(* IEC 61131-3 sources: daoli-st-library/DL_Device (part 9) *)

(* ---- FC_DL_FiberDiameterFromDrawRateCalc.st ---- *)
// FC_DL_FiberDiameterFromDrawRateCalc v1.0.0
// 开源溯源：clean-room 自研（族 DL_Device，ST 生态实测 0 命中，无外部代码引入）
(*
  功能: 由单孔质量流量与拉丝速度反算纤维直径：质量流量 g/h→kg/h→kg/s（除 1000、除 3600），
        除 ρ 得体积流量 [m³/s]，除以 m/s 得截面积 A [m²]，d = 2·SQRT(A/π)·1e6 [µm]。
        注：派单式原写 (m/1000/ρ)/(v/60)，缺 h→s 的 3600 换算；不补则结果恒放大 3600 倍
        （30 g/h、900 m/min、2500 kg/m³ 时得 1009 µm 而非 16.8 µm），3~30 µm 工艺窗永久不可达。
        本件按量纲一致性显式补入 3600，公式其余部分不变。
  邻件/码位: 与 FC_DL_BushingDwellFlowCalc 正串联（前件出单孔流量）；
             16#0002_9223 = 非有限、拉丝速度/密度非正、流量非正或直径出 3~30 µm。
*)
FUNCTION FC_DL_FiberDiameterFromDrawRateCalc : REAL
VAR_INPUT
    fFlowRate  : REAL := 30.0;      // 单孔质量流量 [g/h]，域 > 0 / Mass flow per orifice [g/h]
    fDrawSpeed : REAL := 900.0;     // 拉丝线速度 [m/min]，域 > 0 / Drawing speed [m/min]
    fDensity   : REAL := 2500.0;    // 玻璃密度 [kg/m³]，域 > 0 / Glass density [kg/m^3]
END_VAR
VAR_OUTPUT
    fDiameterUm : REAL;             // 纤维直径 [µm]，工艺窗 3~30 / Fiber diameter [um]
    bValid      : BOOL;             // 结果有效回执 [-] / Result validity receipt
    uErrorId    : UDINT;            // 事件码，0 = 无事件 / Event code
END_VAR
VAR
    fMassKgS : REAL := 0.0;         // 单孔质量流量 [kg/s] / Mass flow [kg/s]
    fVolRate : REAL := 0.0;         // 单孔体积流量 [m³/s] / Volumetric flow [m^3/s]
    fVelocity : REAL := 0.0;        // 拉丝线速度 [m/s] / Drawing speed [m/s]
    fArea    : REAL := 0.0;         // 单丝截面积 [m²] / Filament cross-section [m^2]
END_VAR
// 段 0：全路径出口安全缺省 / Safe defaults on all outlets
fDiameterUm := 0.0;                 // 直径缺省零 / Diameter default zero
bValid := FALSE;                    // 有效回执预清 / Validity preset clear
uErrorId := 16#0000;                // 事件码预清 / Event code preset clear
FC_DL_FiberDiameterFromDrawRateCalc := 0.0; // 返回值缺省零（镜像直径）/ Return default zero
// 段 1：非有限闸（三入参全枚举）/ Non-finite gate over all inputs
IF (fFlowRate <> fFlowRate) OR (fDrawSpeed <> fDrawSpeed) OR (fDensity <> fDensity)
   OR (ABS(fFlowRate) >= 3.0E38) OR (ABS(fDrawSpeed) >= 3.0E38) OR (ABS(fDensity) >= 3.0E38) THEN
    uErrorId := 16#0002_9223;   // 入参非有限拒收 / Non-finite input reject
    RETURN;
END_IF
// 段 2：域闸（拉丝速度与密度为正防除零 + 流量为正，R4）/ Domain gate
IF (fDrawSpeed <= 1.0E-6) OR (fDensity <= 1.0E-6) THEN
    uErrorId := 16#0002_9223;   // 拉丝速度或密度非正 / Non-positive speed or density
    RETURN;
END_IF
IF fFlowRate <= 1.0E-6 THEN
    uErrorId := 16#0002_9223;   // 流量非正（无丝可拉）/ Non-positive flow, no filament
    RETURN;
END_IF
// 段 3：主计算（质量→体积流量→截面积→直径）/ Main computation
fMassKgS := fFlowRate / 1000.0 / 3600.0;                        // 质量流量 [kg/s] / Mass flow
fVolRate := fMassKgS / fDensity;                                // 体积流量 [m³/s] / Volumetric flow
fVelocity := fDrawSpeed / 60.0;                                 // 线速度 [m/s] / Drawing speed
fArea := fVolRate / fVelocity;                                  // 截面积 [m²] / Cross-section area
fDiameterUm := 2.0 * SQRT(fArea / 3.14159265358979) * 1.0E6;    // d = 2·sqrt(A/π) [µm] / Diameter
// 段 4：出口闸（非有限复核 + 3~30 µm 工艺窗判定）/ Outlet gate
IF (fDiameterUm <> fDiameterUm) OR (ABS(fDiameterUm) >= 3.0E38) THEN
    fDiameterUm := 0.0;         // 复核失败回缺省 / Fallback on recheck failure
    uErrorId := 16#0002_9223;   // 出口非有限拒收 / Output non-finite reject
    RETURN;
END_IF
IF (fDiameterUm < 3.0) OR (fDiameterUm > 30.0) THEN
    uErrorId := 16#0002_9223;   // 信息级：直径出 3~30 µm 工艺窗 / Info: diameter out of window
    RETURN;                     // bValid 保持 FALSE / Validity stays false
END_IF
bValid := TRUE;                 // 有效回执 / Validity receipt
FC_DL_FiberDiameterFromDrawRateCalc := fDiameterUm;     // 返回值镜像直径 / Return mirrors diameter
END_FUNCTION

(* ---- FC_DL_ForkEntryClearanceCalc.st ---- *)
(*
  DL Factory R83 | FC_DL_ForkEntryClearanceCalc
  功能：按货位内宽、托盘宽与对中偏差算入叉左右余量，并判叉体能否进槽。
  开源溯源：无（clean-room 自研，依据公开工艺公式，来源=行业通用公式，许可证=MIT，借鉴点=公式结构）
  规则：R1-R21 全遵守
*)
FUNCTION FC_DL_ForkEntryClearanceCalc : REAL
VAR_INPUT
    fSlotWidMm   : REAL; // 货位立柱内侧净宽 [mm] / Slot clear width between uprights [mm]
    fPalletWidMm : REAL; // 托盘宽度 [mm] / Pallet width [mm]
    fForkWidMm   : REAL; // 货叉外廓总宽 [mm] / Fork overall width [mm]
    fOffsetMm    : REAL; // 堆垛机对中偏差（正=偏右）[mm] / Centring offset, + = right [mm]
END_VAR
VAR_OUTPUT
    fLeftMm     : REAL; // 左侧余量 [mm] / Left clearance [mm]
    fRightMm    : REAL; // 右侧余量 [mm] / Right clearance [mm]
    fMinClearMm : REAL; // 双侧最小余量（决定能否入叉）[mm] / Governing minimum clearance [mm]
    xOk         : BOOL; // 入叉判定（最小余量不低于 25 mm）/ Entry decision, at least 25 mm
    xValid      : BOOL; // 计算有效性标志 / Calculation validity flag
END_VAR
VAR
    fGovernWidMm : REAL; // 实际占宽（托盘宽与叉宽取大者）[mm] / Governing occupied width [mm]
    fHalfGapMm   : REAL; // 名义单侧余量 [mm] / Nominal per-side clearance [mm]
END_VAR
fLeftMm := 0.0; fRightMm := 0.0; fMinClearMm := 0.0; xOk := FALSE; xValid := FALSE; // 出口预置
// 非有限拦截 + 量纲自检（R20/R21）
IF NOT (fSlotWidMm > -1.0E30 AND fSlotWidMm < 1.0E30) OR NOT (fPalletWidMm > -1.0E30 AND fPalletWidMm < 1.0E30) OR NOT (fForkWidMm > -1.0E30 AND fForkWidMm < 1.0E30) OR NOT (fOffsetMm > -1.0E30 AND fOffsetMm < 1.0E30) OR fSlotWidMm <= 0.0 OR fPalletWidMm <= 0.0 OR fForkWidMm <= 0.0 THEN
    FC_DL_ForkEntryClearanceCalc := -1.0; RETURN;  // 哨兵 -1：非有限或量纲越界 / Sentinel -1
END_IF
// 实际占宽：托盘与叉体取大者（叉宽超托盘时由叉体决定余量）
IF fPalletWidMm >= fForkWidMm THEN
    fGovernWidMm := fPalletWidMm;   // 托盘占宽为主 [mm] / Pallet governs
ELSE
    fGovernWidMm := fForkWidMm;     // 叉体占宽为主 [mm] / Fork governs
END_IF
// 名义单侧余量：(净宽 - 占宽) ÷ 2，负值表示物理上装不进去
fHalfGapMm := (fSlotWidMm - fGovernWidMm) / 2.0; // 名义单侧余量 [mm] / Nominal per-side clearance
// 左右余量：对中偏差按正负拆分，同量纲（mm）加减，分解后之和恒等于 2×名义余量
fLeftMm  := fHalfGapMm - fOffsetMm;   // 左余量 [mm]，偏右时变小 / Left clearance [mm]
fRightMm := fHalfGapMm + fOffsetMm;   // 右余量 [mm]，偏右时变大 / Right clearance [mm]
// 双侧最小余量：决定可否入叉的瓶颈侧
IF fLeftMm <= fRightMm THEN
    fMinClearMm := fLeftMm;         // 左侧为瓶颈 [mm] / Left is governing
ELSE
    fMinClearMm := fRightMm;        // 右侧为瓶颈 [mm] / Right is governing
END_IF
// 入叉判定：最小余量不低于 25 mm（AGV/堆垛机通用安全余量）
xOk    := fMinClearMm >= 25.0;      // 入叉布尔 / Entry boolean
xValid := TRUE; FC_DL_ForkEntryClearanceCalc := fMinClearMm; // 返回最小余量 [mm] / Return clearance
END_FUNCTION

(* ---- FC_DL_FreeCoolingHoursCalc.st ---- *)
(*
 * FC_DL_FreeCoolingHoursCalc | C2 | DL_Device
 * 功能：逐时干球温度法统计自然冷却可用小时数（含滞环）       单位：温度 [℃]、滞环 [K]、小时 [h]、格数 [1]
 * 工况边界：固定 24 格逐时数组（禁变长数组），每格代表 1 h；判据 outdoor < return − hyst；任一小时数据 NaN/±Inf 或超量程即判 xValid=FALSE 并把可用小时数与最低温度置安全值 0；本件为温度法简化，工程定案须用焓差法复核
 * 代数值回代：return=30 ℃、hyst=2 K → 阈值 28 ℃；若 24 格中 10 格 <28 ℃ → 可用 10 h、nFreeBins=10、rMinOutdoorC=各格最小值（与 spec 1 h/格计数一致）
 * 开源溯源：clean-room 自研，未复制任何第三方代码（无外部来源）
 *)
FUNCTION FC_DL_FreeCoolingHoursCalc : BOOL
VAR_INPUT
    arOutdoorC : ARRAY[1..24] OF REAL;  // 逐时户外干球温度 | hourly outdoor dry bulb temperature [℃]
    rReturnC   : REAL := 30.0;          // 机房回风温度 | room return air temperature [℃]
    rHystK     : REAL := 2.0;           // 自然冷却投入滞环 | free cooling hysteresis [K]
END_VAR
VAR_OUTPUT
    rFreeHours  : REAL;                 // 自然冷却可用小时数 | free cooling available hours [h]
    nFreeBins   : INT;                  // 可用小时格数 | number of free cooling bins [格]
    rMinOutdoorC: REAL;                 // 全年最低户外温度（诊断用）| minimum outdoor temperature for diagnostics [℃]
    xValid      : BOOL;                 // 输出有效 | outputs valid
END_VAR
VAR
    nIdx      : INT;                    // 数组下标 | array index [1]
    nBadBins  : INT;                    // 非法数据格数 | count of non-finite or out-of-range bins [格]
    xFinRet   : BOOL;                   // 回风温度有限性 | return temperature is finite
    xFinHyst  : BOOL;                   // 滞环有限性 | hysteresis is finite
    xBinFin   : BOOL;                   // 单格有限性 | this bin is finite
    rThreshC  : REAL;                   // 自然冷却投入阈值 | free cooling threshold temperature [℃]
    rValC     : REAL;                   // 当前格温度 | current bin temperature [℃]
END_VAR
VAR CONSTANT
    DL_FCH_TEMP_MAX : REAL := 60.0;     // 温度量程上限 | upper temperature limit [℃]
    DL_FCH_TEMP_MIN : REAL := -60.0;    // 温度量程下限 | lower temperature limit [℃]
    DL_FCH_HOUR_PER_BIN : REAL := 1.0;  // 每格代表小时数 | hours represented by one bin [h]
END_VAR

// 段1｜非有限闸：回风温度与滞环（R19）
xFinRet := (rReturnC = rReturnC) AND ((rReturnC - rReturnC) = 0.0);
xFinHyst := (rHystK = rHystK) AND ((rHystK - rHystK) = 0.0);
IF (NOT xFinRet) OR (NOT xFinHyst) OR (rHystK < 0.0) THEN
    rFreeHours := 0.0;                  // 安全值：可用小时 0 | safe value, zero hours
    nFreeBins := 0;
    rMinOutdoorC := 0.0;
    xValid := FALSE;
    FC_DL_FreeCoolingHoursCalc := FALSE;
    RETURN;
END_IF

// 段2｜逐格统计（禁变长数组，固定 1..24）
rThreshC := rReturnC - rHystK;
nFreeBins := 0;
nBadBins := 0;
rMinOutdoorC := arOutdoorC[1];          // 以首格初始化，后续逐格比较 | initialised with the first bin
FOR nIdx := 1 TO 24 DO
    rValC := arOutdoorC[nIdx];
    xBinFin := (rValC = rValC) AND ((rValC - rValC) = 0.0);
    IF (NOT xBinFin) OR (rValC > DL_FCH_TEMP_MAX) OR (rValC < DL_FCH_TEMP_MIN) THEN
        nBadBins := nBadBins + 1;       // 非法格不计入可用，也不参与最低值 | invalid bins are excluded from both statistics
    ELSE
        IF rValC < rThreshC THEN
            nFreeBins := nFreeBins + 1; // 该格计入可用小时 | this bin counts as free cooling time
        END_IF
        IF rValC < rMinOutdoorC THEN
            rMinOutdoorC := rValC;      // 追踪最低温度 | track the minimum
        END_IF
    END_IF
END_FOR

// 段3｜结果：任一杯坏数据即整表判无效（不发布半可信统计）
IF nBadBins > 0 THEN
    rFreeHours := 0.0;                  // 安全值：可用小时 0 | safe value, zero hours
    nFreeBins := 0;
    rMinOutdoorC := 0.0;
    xValid := FALSE;
    FC_DL_FreeCoolingHoursCalc := FALSE;
    RETURN;
END_IF
rFreeHours := INT_TO_REAL(nFreeBins) * DL_FCH_HOUR_PER_BIN;

// 段4｜出口
xValid := TRUE;
FC_DL_FreeCoolingHoursCalc := TRUE;
END_FUNCTION

(* ---- FC_DL_HydroAccumulatorSizing.st ---- *)
(*
  ============================================================
  组件名 : FC_DL_HydroAccumulatorSizing
  分类   : DL_Device
  功能   : 皮囊式蓄能器容积选型，按等温或绝热过程由需液量、最高最低压力与预充压力求公称容积
  开源溯源 : internal-design（本轮无外部代码逐行引用）
             参考语义 : 无外部参考
  复杂度 : C2
  版本   : 1.0.0
  ============================================================
*)

FUNCTION FC_DL_HydroAccumulatorSizing : REAL
VAR_INPUT
    rVolumeDemand_l    : REAL; // 需液量 [l] usable oil demand [litre]
    rPressMax_bar      : REAL; // 最高工作压力 [bar] maximum working pressure [bar]
    rPressMin_bar      : REAL; // 最低工作压力 [bar] minimum working pressure [bar]
    rPressPrecharge_bar: REAL; // 预充压力 [bar] precharge pressure [bar]
    bAdiabatic         : BOOL; // 真为绝热过程，假为等温过程 adiabatic when true, isothermal when false
END_VAR
VAR_OUTPUT
    rVolume_l     : REAL; // 蓄能器公称容积 [l] nominal accumulator volume [litre]
    rUsableRatio  : REAL; // 有效容积比 [无量纲] usable volume ratio [dimensionless]
    bValid        : BOOL; // 结果有效标志 result validity flag
END_VAR
VAR CONSTANT
    DL_ADIA_EXP : REAL := 0.7142857; // 绝热指数倒数值 1/1.4 reciprocal of the adiabatic index
    DL_EPS_R    : REAL := 1.0E-6; // 实数零判定阈值 real zero threshold
END_VAR
VAR
    _bFin   : BOOL := FALSE; // 四实数输入有限性判定 finiteness verdict of the four real inputs
    _rRatio : REAL := 0.0; // 压比 the pressure ratio [dimensionless]
    _rProc  : REAL := 0.0; // 过程指数折算后的压比 the process weighted pressure ratio [dimensionless]
    _rDen   : REAL := 0.0; // 容积公式分母 [无量纲] denominator of the volume formula [dimensionless]
    _rVol   : REAL := 0.0; // 公称容积中间量 [l] intermediate nominal volume [litre]
END_VAR

// 段 1｜出口预置 preset the exit
FC_DL_HydroAccumulatorSizing := 0.0; // 缺省返回零 default zero return
rVolume_l := 0.0; // 容积预置零 volume preset to zero
rUsableRatio := 0.0; // 有效容积比预置零 usable ratio preset to zero
bValid := FALSE; // 计算完成前不认结果 unusable before the calculation
// 段 2｜非有限闸 finiteness gate
_bFin := (rVolumeDemand_l = rVolumeDemand_l) AND (rPressMax_bar = rPressMax_bar) AND (rPressMin_bar = rPressMin_bar) AND (rPressPrecharge_bar = rPressPrecharge_bar); // 四输入自反判定 self comparison of the four inputs
IF NOT _bFin THEN
    RETURN; // 非有限即无效 non finite means invalid
END_IF
// 段 3｜压力几何闸 pressure geometry gate
IF rPressMin_bar <= 0.0 THEN
    RETURN; // 最低压力非正无法形成压比 a non positive minimum cannot form a ratio
END_IF
IF (rPressMax_bar <= rPressMin_bar) OR (rPressMin_bar <= rPressPrecharge_bar) THEN
    RETURN; // 高压须大于低压，低压须大于预充 the maximum must exceed the minimum and the minimum must exceed the precharge
END_IF
IF rVolumeDemand_l < 0.0 THEN
    RETURN; // 需液量为负属配置非法 a negative demand is an illegal configuration
END_IF
// 段 4｜过程折算与分母 process weighting and the denominator
_rRatio := rPressMax_bar / rPressMin_bar; // 最高与最低压力比 ratio of the maximum to the minimum
IF bAdiabatic THEN
    _rProc := EXPT(_rRatio, DL_ADIA_EXP); // 绝热过程按一点四指数折算 adiabatic process weighted by the index of one point four
ELSE
    _rProc := _rRatio; // 等温过程压比直通 isothermal process keeps the plain ratio
END_IF
_rDen := _rProc - 1.0; // 容积公式分母 denominator of the volume formula
IF _rDen <= DL_EPS_R THEN
    RETURN; // 分母近零无法定容 a near zero denominator cannot size the volume
END_IF
// 段 5｜公称容积与有效容积比 nominal volume and the usable ratio
_rVol := rVolumeDemand_l / _rDen; // 公称容积 nominal volume
rVolume_l := _rVol; // 容积落定 land the volume
rUsableRatio := rVolumeDemand_l / _rVol; // 有效容积比 usable volume ratio
bValid := TRUE; // 结果可用 result usable
FC_DL_HydroAccumulatorSizing := _rVol; // 函数返回公称容积 return the nominal volume
END_FUNCTION

(* ---- FC_DL_HydroCylFlowNeed.st ---- *)
(*
  ============================================================
  组件名 : FC_DL_HydroCylFlowNeed
  分类   : DL_Device
  功能   : 液压缸动作所需流量计算，由有效面积、目标速度与容积效率求泵侧流量
  开源溯源 : internal-design（本轮无外部代码逐行引用）
             参考语义 : 无外部参考
  复杂度 : C1
  版本   : 1.0.0
  ============================================================
*)

FUNCTION FC_DL_HydroCylFlowNeed : REAL
VAR_INPUT
    rArea_cm2  : REAL; // 有效作用面积 [cm2] effective acting area [cm2]
    rSpeed_mm_s: REAL; // 目标速度 [mm/s] target speed [mm per second]
    rVolEff    : REAL; // 容积效率 0~1 [无量纲] volumetric efficiency from zero to one [dimensionless]
END_VAR
VAR_OUTPUT
    rFlow_lpm : REAL; // 所需流量 [l/min] required flow [litre per minute]
    bValid    : BOOL; // 结果有效标志 result validity flag
END_VAR
VAR CONSTANT
    DL_MM_PER_CM    : REAL := 10.0; // 每厘米毫米数 millimetres per centimetre
    DL_SEC_PER_MIN  : REAL := 60.0; // 每分钟秒数 seconds per minute
    DL_CM3_PER_L    : REAL := 1000.0; // 每升立方厘米数 cubic centimetres per litre
END_VAR
VAR
    _bFin  : BOOL := FALSE; // 三输入有限性判定 finiteness verdict of the three inputs
    _rVelCms : REAL := 0.0; // 速度折算 [cm/s] speed in centimetres per second [cm/s]
    _rFlow : REAL := 0.0; // 流量中间量 [l/min] intermediate flow [litre per minute]
END_VAR

// 段 1｜出口预置 preset the exit
FC_DL_HydroCylFlowNeed := 0.0; // 缺省返回零 default zero return
rFlow_lpm := 0.0; // 流量预置零 flow preset to zero
bValid := FALSE; // 计算完成前不认结果 unusable before the calculation
// 段 2｜非有限闸 finiteness gate
_bFin := (rArea_cm2 = rArea_cm2) AND (rSpeed_mm_s = rSpeed_mm_s) AND (rVolEff = rVolEff); // 三输入自反判定 self comparison of the three inputs
IF NOT _bFin THEN
    RETURN; // 非有限即无效 non finite means invalid
END_IF
// 段 3｜面积与效率闸 area and efficiency gate
IF (rArea_cm2 <= 0.0) OR (rSpeed_mm_s < 0.0) THEN
    RETURN; // 面积非正或负速度属配置非法 an illegal area or a negative speed
END_IF
IF (rVolEff <= 0.0) OR (rVolEff > 1.0) THEN
    RETURN; // 容积效率越出零到一 volumetric efficiency outside the open closed interval
END_IF
// 段 4｜主体换算 main unit conversion
_rVelCms := rSpeed_mm_s / DL_MM_PER_CM; // 毫米每秒折算为厘米每秒 convert millimetres to centimetres per second
_rFlow := rArea_cm2 * _rVelCms * DL_SEC_PER_MIN / DL_CM3_PER_L; // 面积乘速度得流量 area times speed gives the flow
_rFlow := _rFlow / rVolEff; // 容积效率折损修正 volumetric loss correction
rFlow_lpm := _rFlow; // 流量落定 land the flow
bValid := TRUE; // 结果可用 result usable
FC_DL_HydroCylFlowNeed := _rFlow; // 函数返回流量 return the flow
END_FUNCTION

(* ---- FC_DL_HydroCylForceCalc.st ---- *)
(*
  ============================================================
  组件名 : FC_DL_HydroCylForceCalc
  分类   : DL_Device
  功能   : 液压缸理论推力计算，按缸径杆径、供油压力、背压与机械效率求伸出与缩回推力
  开源溯源 : internal-design（本轮无外部代码逐行引用）
             参考语义 : 无外部参考
  复杂度 : C1
  版本   : 1.0.0
  ============================================================
*)

FUNCTION FC_DL_HydroCylForceCalc : REAL
VAR_INPUT
    rBoreDia_mm  : REAL; // 缸径 [mm] bore diameter [mm]
    rRodDia_mm   : REAL; // 活塞杆径 [mm] rod diameter [mm]
    rPressBar    : REAL; // 供油压力 [bar] supply pressure [bar]
    rBackPressBar: REAL; // 回油背压 [bar] return line back pressure [bar]
    rMechEff     : REAL; // 机械效率 0~1 [无量纲] mechanical efficiency from zero to one [dimensionless]
    bExtend      : BOOL; // 真为伸出，假为缩回 extend when true, retract when false
END_VAR
VAR_OUTPUT
    rForce_kN : REAL; // 理论推力 [kN] theoretical force [kN]
    rArea_cm2 : REAL; // 有效作用面积 [cm2] effective acting area [cm2]
    bValid    : BOOL; // 结果有效标志 result validity flag
END_VAR
VAR CONSTANT
    DL_PI_4     : REAL := 0.7853982; // 四分之圆周率 pi divided by four
    DL_MM2_PER_CM2 : REAL := 100.0; // 平方毫米到平方厘米换算 square millimetres per square centimetre
    DL_BAR_TO_KPA : REAL := 100.0; // 巴到千帕换算 kilopascal per bar
END_VAR
VAR
    _bFin   : BOOL := FALSE; // 五实数输入有限性判定 finiteness verdict of the five real inputs
    _rAreaMM2 : REAL := 0.0; // 有效面积 [mm2] effective area [mm2]
    _rDpBar : REAL := 0.0; // 有效压差 [bar] effective pressure difference [bar]
    _rForce : REAL := 0.0; // 推力中间量 [kN] intermediate force [kN]
END_VAR

// 段 1｜出口预置 preset the exit
FC_DL_HydroCylForceCalc := 0.0; // 缺省返回零 default zero return
rForce_kN := 0.0; // 推力预置零 force preset to zero
rArea_cm2 := 0.0; // 面积预置零 area preset to zero
bValid := FALSE; // 计算完成前不认结果 unusable before the calculation
// 段 2｜非有限闸 finiteness gate
_bFin := (rBoreDia_mm = rBoreDia_mm) AND (rRodDia_mm = rRodDia_mm) AND (rPressBar = rPressBar) AND (rBackPressBar = rBackPressBar) AND (rMechEff = rMechEff); // 五输入自反判定 self comparison of the five inputs
IF NOT _bFin THEN
    RETURN; // 非有限即无效 non finite means invalid
END_IF
// 段 3｜几何与效率闸 geometry and efficiency gate
IF (rBoreDia_mm <= 0.0) OR (rRodDia_mm < 0.0) THEN
    RETURN; // 缸径非正或杆径为负属配置非法 an illegal bore or rod geometry
END_IF
IF (rMechEff <= 0.0) OR (rMechEff > 1.0) THEN
    RETURN; // 效率越出零到一 efficiency outside the open closed interval
END_IF
IF (rPressBar < 0.0) OR (rBackPressBar < 0.0) THEN
    RETURN; // 负压力属配置非法 a negative pressure is an illegal configuration
END_IF
// 段 4｜有效面积：伸出取缸径面积，缩回取环形面积 effective area of both directions
IF bExtend THEN
    _rAreaMM2 := DL_PI_4 * rBoreDia_mm * rBoreDia_mm; // 缸径全截面 full bore section
ELSE
    IF (rRodDia_mm <= 0.0) OR (rRodDia_mm >= rBoreDia_mm) THEN
        RETURN; // 缩回要求杆径在零与缸径之间 retraction needs a rod between zero and the bore
    END_IF
    _rAreaMM2 := DL_PI_4 * (rBoreDia_mm * rBoreDia_mm - rRodDia_mm * rRodDia_mm); // 环形截面 annulus section
END_IF
rArea_cm2 := _rAreaMM2 / DL_MM2_PER_CM2; // 面积换算为平方厘米 convert the area to square centimetres
// 段 5｜压差与推力 pressure difference and the force
_rDpBar := rPressBar - rBackPressBar; // 有效压差 effective pressure difference
_rForce := _rDpBar * DL_BAR_TO_KPA * rArea_cm2 / 10000.0 * rMechEff; // 千帕乘平方米得千牛 kilopascal times square metre gives kilonewton
rForce_kN := _rForce; // 推力落定 land the force
bValid := TRUE; // 结果可用 result usable
FC_DL_HydroCylForceCalc := _rForce; // 函数返回推力 return the force
END_FUNCTION

(* ---- FC_DL_InventoryAgeIndexCalc.st ---- *)
(*
  DL Factory R83 | FC_DL_InventoryAgeIndexCalc
  功能：把库龄与周转等级加权成 0~100 出库优先级指数，并给出优先级别与判定。
  开源溯源：无（clean-room 自研，依据公开工艺公式，来源=行业通用公式，许可证=MIT，借鉴点=公式结构）
  规则：R1-R21 全遵守
*)
FUNCTION FC_DL_InventoryAgeIndexCalc : REAL
VAR_INPUT
    fAgeDays    : REAL; // 当前库龄 [天] / Current inventory age [days]
    fMaxAgeDays : REAL; // 库龄归一化上限（超过按满分）[天] / Age normalisation ceiling [days]
    iTurnClass  : INT;  // 周转等级 1=快 2=中 3=慢 / Turnover class 1=fast 2=medium 3=slow
    fWeightAge  : REAL; // 库龄权重（0~1，其余给周转等级）[-]/ Age weight, remainder to turnover [-]
END_VAR
VAR_OUTPUT
    fAgeScore : REAL; // 库龄得分（0~100）[-]/ Age score [0..100]
    fAgeIdx   : REAL; // 综合库龄指数（0~100）[-]/ Composite age index [0..100]
    iPrioLvl  : INT;  // 优先级别 1=最高 2=中 3=低 / Priority level 1=highest 3=lowest
    xPriority : BOOL; // 优先出库判定（指数不低于 60）/ Priority pick flag, index at or above 60
    xValid    : BOOL; // 计算有效性标志 / Calculation validity flag
END_VAR
VAR
    fTurnScore : REAL; // 周转等级得分（0~100）[-]/ Turnover score [0..100]
END_VAR
// 出口预置：五出口统一预置，优先级默认最低（安全侧）
fAgeScore := 0.0; fAgeIdx := 0.0; iPrioLvl := 3; xPriority := FALSE; xValid := FALSE;
// 非有限拦截 + 量纲自检 + 周转等级域闸（R20/R21）
IF NOT (fAgeDays > -1.0E30 AND fAgeDays < 1.0E30) OR NOT (fMaxAgeDays > -1.0E30 AND fMaxAgeDays < 1.0E30) OR NOT (fWeightAge > -1.0E30 AND fWeightAge < 1.0E30) OR fAgeDays < 0.0 OR fMaxAgeDays <= 0.0 OR iTurnClass < 1 OR iTurnClass > 3 OR fWeightAge < 0.0 OR fWeightAge > 1.0 THEN
    FC_DL_InventoryAgeIndexCalc := -1.0; RETURN; // 哨兵 -1：非有限或量纲/等级越界 / Sentinel -1
END_IF
// 库龄得分：库龄 ÷ 上限 × 100；超上限先判并封顶 100，避免饱和逻辑与实数上限冲突（R28）
IF fAgeDays >= fMaxAgeDays THEN
    fAgeScore := 100.0;             // 达到归一化上限，满分 / At ceiling, full score
ELSE
    fAgeScore := (fAgeDays / fMaxAgeDays) * 100.0;  // 线性归一化得分 / Linear normalised score
END_IF
// 周转等级得分：等级 1→100，2→66.7，3→33.3，即 (4 - 等级) ÷ 3 × 100
fTurnScore := (INT_TO_REAL(4 - iTurnClass) / 3.0) * 100.0;  // 周转得分 [-] / Turnover score
// 综合指数：库龄权重 × 库龄得分 + (1 - 权重) × 周转得分，权重和为 1 故仍 0~100
fAgeIdx := fWeightAge * fAgeScore + (1.0 - fWeightAge) * fTurnScore; // 综合指数 [-] / Composite index
// 优先级分档：指数越高越先出库，分界 80 / 60（严格不等，禁浮点等号）
IF fAgeIdx >= 80.0 THEN
    iPrioLvl := 1;                  // 最高优先级 / Highest priority
ELSIF fAgeIdx >= 60.0 THEN
    iPrioLvl := 2;                  // 中优先级 / Medium priority
ELSE
    iPrioLvl := 3;                  // 低优先级 / Low priority
END_IF
xPriority := fAgeIdx >= 60.0;       // 优先出库判定 / Priority pick flag
xValid := TRUE; FC_DL_InventoryAgeIndexCalc := fAgeIdx;  // 链路有效并返回综合指数 [-]
END_FUNCTION

(* ---- FC_DL_KcellConstCalc.st ---- *)
(* ============================================================
   DL_Device / FC_DL_KcellConstCalc ｜ v1.0.0 ｜ 2026-11-25
   功能：电导池常数标定反算 Kcell = σ_std · R_meas [1/cm]（σ 由 µS/cm ×1E-6 转 S/cm），
         温度修正 K_tcorr = Kcell / (1 + α·(T − 25))，α = fTempCoefPct / 100。
   边界：标准液电导率 ≤ 0 或实测电阻 ≤ 0 → 两出口写 0、码 1（N1：值与判据同拍改写）；
         任一入参非有限 → 两出口写 0、码 2；温补分母 ≤ 0.01 → 码 3 且温度修正值
         回退为未修正值（不给伪修正结果）。
         量纲清单（N5）：1 S/cm = 1E6 µS/cm；1 Ω⁻¹ = 1 S；Kcell 单位 1/cm；
         回代：σ=1413 µS/cm、R=100 Ω → 0.1413 1/cm。
   依赖：仅 IEC 61131-3（无外部依赖，纯算术） ｜ 溯源：DLF-D-WATERANA
   验收：1413 µS/cm、100 Ω → Kcell=0.1413 1/cm、码 0；T=35、α=2%/°C →
         K_tcorr = 0.1413 / 1.2 = 0.1178 1/cm；σ=0 → 码 1、两出口 0。
   ============================================================ *)
FUNCTION FC_DL_KcellConstCalc : BOOL
VAR_INPUT
    fStdUsCm     : REAL;  // 标准液电导率（25°C 标称值）[µS/cm] / Conductivity of the standard solution
    fRMeasOhm    : REAL;  // 实测电导池电阻 [Ω] / Measured conductivity cell resistance
    fTempC       : REAL;  // 标准液实测温度 [°C] / Measured temperature of the standard solution
    fTempCoefPct : REAL;  // 电导率温补系数（%/°C，常取 2.0）[%/°C] / Conductivity temperature coefficient
END_VAR
VAR_OUTPUT
    fKcell      : REAL;   // 未温度修正的池常数 [1/cm] / Cell constant without temperature correction
    fKcellTcorr : REAL;   // 温度修正后池常数 [1/cm] / Temperature corrected cell constant
    uErrId      : UDINT;  // 码 0 正常 / 1 域闸 / 2 非有限 / 3 温补分母非法 [-] / Outlet code
END_VAR
VAR
    _fK     : REAL;  // 未修正池常数中间值 [1/cm] / Intermediate uncorrected cell constant
    _fDen   : REAL;  // 温补分母 (1 + α·(T−25)) [-] / Temperature correction denominator
    _bDen   : BOOL;  // 温补分母非法标志 [-] / Illegal denominator flag
END_VAR
VAR CONSTANT
    DL_KCL_US_TO_S : REAL := 1.0E-6;  // µS/cm → S/cm 换算系数 [S·cm/µS] / Microsiemens per centimeter to siemens per centimeter
    DL_KCL_TREF    : REAL := 25.0;    // 参考温度 [°C] / Reference temperature
    DL_KCL_HUND    : REAL := 100.0;   // 百分比换算系数 [%] / Percent conversion factor
    DL_KCL_DFLOOR  : REAL := 0.01;    // 温补分母下限 [-] / Lower bound of the temperature denominator
    DL_KCL_DCEIL   : REAL := 10.0;    // 温补分母上限（防分母虚高致池常数偏低）[-] / Upper bound of the temperature denominator
END_VAR

(* 段 0：出口预置安全侧（两出口 0、码取最严，N1/N3） *)
FC_DL_KcellConstCalc := FALSE;
fKcell := 0.0;  fKcellTcorr := 0.0;  uErrId := 2;
_bDen := FALSE;

(* 段 1：非有限闸（四个入参全量枚举；NaN 自反 + Inf 差值自减双判，R79/R272） *)
IF (fStdUsCm <> fStdUsCm) OR (fRMeasOhm <> fRMeasOhm)
   OR (fTempC <> fTempC) OR (fTempCoefPct <> fTempCoefPct) THEN RETURN; END_IF
(* Inf 双判须覆盖 fTempC：温度 +Inf 使温补分母为 Inf、修正值算成 0，却报 uErrId=0
   成功（伪有效池常数，下游按 k=0 换算全量程失真） *)
IF ((fStdUsCm - fStdUsCm) <> (fStdUsCm - fStdUsCm))
   OR ((fRMeasOhm - fRMeasOhm) <> (fRMeasOhm - fRMeasOhm))
   OR ((fTempC - fTempC) <> (fTempC - fTempC))
   OR ((fTempCoefPct - fTempCoefPct) <> (fTempCoefPct - fTempCoefPct)) THEN RETURN; END_IF

(* 段 2：域闸（电导率与电阻必须为正，防零与负物理量） *)
IF (fStdUsCm <= 0.0) OR (fRMeasOhm <= 0.0) THEN
    uErrId := 1;                        // 域闸：无池常数可解
    RETURN;
END_IF

(* 段 3：池常数（乘加，无除法） *)
_fK := fStdUsCm * DL_KCL_US_TO_S * fRMeasOhm;
IF (_fK <> _fK) OR ((_fK - _fK) <> (_fK - _fK)) THEN RETURN; END_IF

(* 段 4：温补分母（除子结构判定，不做伪修正） *)
_fDen := 1.0 + (fTempCoefPct / DL_KCL_HUND) * (fTempC - DL_KCL_TREF);
IF (_fDen <= DL_KCL_DFLOOR) OR (_fDen > DL_KCL_DCEIL) THEN _bDen := TRUE; END_IF   // 双端闸：分母过小放大、过大压缩均判非法 / two-sided guard

(* 段 5：单一出口裁决（两出口同源赋值一次，N4/R23） *)
fKcell := _fK;
IF _bDen THEN
    fKcellTcorr := _fK;                 // 分母非法：回退未修正值
    uErrId      := 3;
ELSE
    fKcellTcorr := _fK / _fDen;         // 分母已证 > 0.01
    uErrId      := 0;  FC_DL_KcellConstCalc := TRUE;
END_IF

(* 段 6：出口非有限复检（同族补修：比值溢出同样禁报码 0 成功，N1） *)
IF (fKcell <> fKcell) OR ((fKcell - fKcell) <> (fKcell - fKcell))
   OR (fKcellTcorr <> fKcellTcorr) OR ((fKcellTcorr - fKcellTcorr) <> (fKcellTcorr - fKcellTcorr)) THEN
    fKcell := 0.0;  fKcellTcorr := 0.0;  uErrId := 2;  FC_DL_KcellConstCalc := FALSE;
END_IF
END_FUNCTION

(* ---- FC_DL_KilnSpecificHeatCalc.st ---- *)
(*
  DL Factory R84 | FC_DL_KilnSpecificHeatCalc
  功能：算单位熟料热耗并折算标准煤耗与实物煤耗
  开源溯源：无（clean-room 自研，依据公开工艺公式，来源=行业通用公式，许可证=MIT，借鉴点=公式结构）
  规则：R1-R16 全遵守
*)
FUNCTION FC_DL_KilnSpecificHeatCalc : REAL
VAR_INPUT
    fFuelKgh : REAL := 8000.0; // 燃料消耗量（实物煤） [kg/h] / fuel consumption [kg/h]
    fLhvKcalkg : REAL := 5500.0; // 燃料低位热值 [kcal/kg] / lower heating value [kcal/kg]
    fClinkerTph : REAL := 250.0; // 熟料产量 [t/h] / clinker output [t/h]
    fKgceKcalkg : REAL := 7000.0; // 标准煤当量热值 [kcal/kgce] / standard coal equivalent [kcal/kgce]
END_VAR
VAR_OUTPUT
    fKgcePerT : REAL; // 折标准煤耗 [kgce/t] / standard coal consumption [kgce/t]
    fCoalRate : REAL; // 实物煤耗 [kg/t] / actual coal rate [kg/t]
    xValid : BOOL; // 计算结果有效标志 [-] / calculation valid flag [-]
END_VAR
VAR
    fKcalH : REAL; // 小时供热量 [kcal/h] / hourly heat input [kcal/h]
    fClinkerKgh : REAL; // 熟料小时产量折算 [kg/h] / clinker output in kilograms [kg/h]
    fSpecKcalkg : REAL; // 单位熟料热耗 [kcal/kg] / specific heat consumption [kcal/kg]
END_VAR

// 段 1｜出口预置（R256）
FC_DL_KilnSpecificHeatCalc := -1.0; // 哨兵返回 -1（无效） [-] / sentinel return -1, invalid [-]
fKgcePerT := 0.0; // 标煤耗预置零 [kgce/t] / standard coal preset zero [kgce/t]
fCoalRate := 0.0; // 实物煤耗预置零 [kg/t] / actual coal rate preset zero [kg/t]
xValid := FALSE; // 计算完成前不认结果 [-] / unusable before calculation [-]

// 段 2｜非有限拦截 + 域闸（R4/R20）
IF NOT (fFuelKgh > -1.0E30 AND fFuelKgh < 1.0E30) OR NOT (fLhvKcalkg > -1.0E30 AND fLhvKcalkg < 1.0E30) OR NOT (fClinkerTph > -1.0E30 AND fClinkerTph < 1.0E30) OR NOT (fKgceKcalkg > -1.0E30 AND fKgceKcalkg < 1.0E30) THEN
    RETURN; // 任一入参为 NaN/Inf 一律拒绝 [-] / any NaN or Inf input rejected [-]
END_IF
IF fFuelKgh < 0.0 OR fLhvKcalkg < 1.0E-9 OR fKgceKcalkg < 1.0E-9 THEN
    RETURN; // 热值与标煤当量正域分母闸（防除零） [kcal/kg] / positive denominator gate [kcal/kg]
END_IF
IF fClinkerTph < 1.0E-9 THEN
    RETURN; // 熟料产量正域分母闸（防除零） [t/h] / clinker output denominator gate [t/h]
END_IF

// 段 3｜单位热耗 = 燃料量 × 低位热值 / 熟料产量
fKcalH := fFuelKgh * fLhvKcalkg; // kg/h × kcal/kg = kcal/h / [kg/h] × [kcal/kg] = [kcal/h]
fClinkerKgh := fClinkerTph * 1000.0; // t/h × 1000 kg/t = kg/h / [t/h] × [kg/t] = [kg/h]
fSpecKcalkg := fKcalH / fClinkerKgh; // kcal/h ÷ kg/h = kcal/kg / [kcal/h] / [kg/h] = [kcal/kg]
IF NOT (fSpecKcalkg > -1.0E30 AND fSpecKcalkg < 1.0E30) THEN
    RETURN; // 结果非有限再拦一次 [-] / second finiteness gate [-]
END_IF

// 段 4｜折标煤与实物煤耗
fKgcePerT := (fSpecKcalkg / fKgceKcalkg) * 1000.0; // (kcal/kg ÷ kcal/kgce) × 1000 kg/t = kgce/t / [kcal/kg]/[kcal/kgce]×[kg/t] = [kgce/t]
fCoalRate := fFuelKgh / fClinkerTph; // kg/h ÷ t/h = kg/t / [kg/h] / [t/h] = [kg/t]
IF NOT (fKgcePerT > -1.0E30 AND fKgcePerT < 1.0E30) OR NOT (fCoalRate > -1.0E30 AND fCoalRate < 1.0E30) THEN
    RETURN; // 结果非有限再拦一次 [-] / second finiteness gate on the results [-]
END_IF
xValid := TRUE; // 链路有效 [-] / chain valid [-]
FC_DL_KilnSpecificHeatCalc := fSpecKcalkg; // 返回单位热耗 [kcal/kg] / return the specific heat [kcal/kg]
END_FUNCTION

(* ---- FC_DL_LubeIntervalCalc.st ---- *)
(*
  道莅工业代码库 / Daoli Industrial ST Library
  组件: FC_DL_LubeIntervalCalc
  分类: DL_Device
  开源溯源: 无（clean-room 工程公式自研；参考公开工艺计算公式，未复制任何受版权保护代码）
  许可证: 本项目自有 (MIT)
  功能: 按负荷、温度、粉尘三指数折算润滑间隔（基准除以三因子乘积），含因子与乘积双闸
*)
FUNCTION FC_DL_LubeIntervalCalc : BOOL
VAR_INPUT
    rBaseH : REAL; // 基准润滑间隔 [h] / base lubrication interval
    rLoadIdx : REAL; // 负荷指数 [-]，域 0~1.5 / load index
    rTempIdx : REAL; // 温度指数 [-]，域 0~1.5 / temperature index
    rDustIdx : REAL; // 粉尘指数 [-]，域 0~1.5 / dust index
END_VAR
VAR_OUTPUT
    rIntervalH : REAL; // 折算后润滑间隔 [h] / corrected lubrication interval
    bValid : BOOL; // 结果有效位 [-] / result valid flag
    iErrCode : INT; // 事件码 0=正常 1=基准间隔非法 2=因子乘积过小已钳位 3=结果非有限 / event code
END_VAR
VAR CONSTANT
    rIdxLo : REAL := 0.2; // 单因子钳位下限 [-] / per-factor clamp floor
    rIdxHi : REAL := 2.0; // 单因子钳位上限 [-] / per-factor clamp ceiling
    rProdMin : REAL := 0.1; // 乘积下限，低于此则间隔不可信 [-] / product floor
    rProdFloor : REAL := 0.2; // 乘积过小时的替代值 [-] / substitute product applied when floored
END_VAR
VAR
    rLoadUse : REAL; // 生效负荷因子 [-] / effective load factor
    rTempUse : REAL; // 生效温度因子 [-] / effective temperature factor
    rDustUse : REAL; // 生效粉尘因子 [-] / effective dust factor
    rProd : REAL; // 三因子乘积 [-] / product of factors
    rProdUse : REAL; // 生效乘积 [-] / effective product
    rIntRaw : REAL; // 未校验间隔 [h] / unchecked interval
END_VAR

    // —— 段 0：全路径预清 —— //
    rLoadUse := 1.0;
    rTempUse := 1.0;
    rDustUse := 1.0;
    rProd := 0.0;
    rProdUse := rProdFloor; // 生效乘积缺省取替代值 [-] / effective product defaults to the floor
    rIntRaw := 0.0;
    rIntervalH := 0.0;
    bValid := FALSE;
    iErrCode := 0;
    FC_DL_LubeIntervalCalc := FALSE;
    // —— 段 1：基准间隔域闸（兼最终分母的来源量） —— //
    IF rBaseH <= 0.0 THEN
        iErrCode := 1; // 基准间隔非法，间隔无定义 / invalid base interval
        RETURN;
    END_IF;
    // —— 段 2：三因子各自钳位到 [0.2, 2.0]（配置越界按边界处理，不中断） —— //
    IF rLoadIdx < rIdxLo THEN
        rLoadUse := rIdxLo; // 下限钳位 / clamp low
    ELSIF rLoadIdx > rIdxHi THEN
        rLoadUse := rIdxHi; // 上限钳位 / clamp high
    ELSE
        rLoadUse := rLoadIdx;
    END_IF;
    IF rTempIdx < rIdxLo THEN
        rTempUse := rIdxLo;
    ELSIF rTempIdx > rIdxHi THEN
        rTempUse := rIdxHi;
    ELSE
        rTempUse := rTempIdx;
    END_IF;
    IF rDustIdx < rIdxLo THEN
        rDustUse := rIdxLo;
    ELSIF rDustIdx > rIdxHi THEN
        rDustUse := rIdxHi;
    ELSE
        rDustUse := rDustIdx;
    END_IF;
    // —— 段 3：乘积闸（分母不得过小，否则间隔被无限拉长） —— //
    rProd := rLoadUse * rTempUse * rDustUse; // 三因子乘积 [-] / product
    IF rProd < rProdMin THEN
        rProdUse := rProdFloor; // 取替代常数（0.2），间隔最多放大 5 倍 / substitute product, interval at most 5x
        iErrCode := 2; // 信息级：乘积过小已钳位 / info level: product floored
    ELSE
        rProdUse := rProd;
    END_IF;
    // —— 段 4：量纲链 (h)/((-)×(-)×(-)) = h —— //
    rIntRaw := rBaseH / rProdUse; // 折算间隔 [h] / corrected interval
    IF ABS(rIntRaw) > 1.0E15 THEN
        iErrCode := 3; // 结果非有限，强制归零 / non-finite result, forced to zero
        RETURN;
    END_IF;
    rIntervalH := rIntRaw;
    bValid := TRUE;
    FC_DL_LubeIntervalCalc := TRUE;
END_FUNCTION

(* ---- FC_DL_MtbfCalc.st ---- *)
(*
  道莅工业代码库 / Daoli Industrial ST Library
  组件: FC_DL_MtbfCalc
  分类: DL_Device
  开源溯源: 无（clean-room 工程公式自研；参考公开工艺计算公式，未复制任何受版权保护代码）
  许可证: 本项目自有 (MIT)
  功能: MTBF / MTTR / 可用率计算，含无失效样本的退化口径
*)
FUNCTION FC_DL_MtbfCalc : BOOL
VAR_INPUT
    rRunHours : REAL; // 统计窗内累计运行小时 [h] / accumulated running hours in window
    rFailCount : REAL; // 统计窗内失效次数 [次] / failure count in window
    rRepairHours : REAL; // 统计窗内累计修复停机小时 [h] / accumulated repair downtime
END_VAR
VAR_OUTPUT
    rMtbfH : REAL; // 平均无故障间隔 [h] / mean time between failures
    rMttrH : REAL; // 平均修复时间 [h] / mean time to repair
    rAvailPct : REAL; // 可用率 [%] / availability
    bValid : BOOL; // 结果有效位 [-] / result valid flag
    iErrCode : INT; // 事件码 0=正常 1=失效次数为负 2=无失效样本（MTBF 取运行小时）3=结果非有限 4=运行小时非正 5=修复小时为负 / event code
END_VAR
VAR CONSTANT
    rInvPct : REAL := 100.0; // 可用率百分数系数 [%] / percentage factor
    rAvailCap : REAL := 100.0; // 可用率饱和上限 [%] / availability cap
END_VAR
VAR
    rFailUse : REAL; // 生效失效次数 [次] / effective failure count
    rMtbfRaw : REAL; // 未校验 MTBF [h] / unchecked MTBF
    rMttrRaw : REAL; // 未校验 MTTR [h] / unchecked MTTR
    rDenom : REAL; // 可用率分母 [h] / availability denominator
END_VAR

    // —— 段 0：全路径预清 —— //
    rFailUse := 0.0;
    rMtbfRaw := 0.0;
    rMttrRaw := 0.0;
    rDenom := 0.0;
    rMtbfH := 0.0;
    rMttrH := 0.0;
    rAvailPct := 0.0;
    bValid := FALSE;
    iErrCode := 0;
    FC_DL_MtbfCalc := FALSE;
    // —— 段 1：失效次数域闸 —— //
    IF rFailCount < 0.0 THEN
        iErrCode := 1; // 失效次数为负，统计口径非法 / negative failure count
        RETURN;
    END_IF;
    IF rRunHours <= 0.0 THEN
        iErrCode := 4; // 运行小时非正，MTBF 无定义 / non-positive running hours
        RETURN;
    END_IF;
    IF rRepairHours < 0.0 THEN
        iErrCode := 5; // 修复小时为负，统计口径非法 / negative repair hours
        RETURN;
    END_IF;
    // —— 段 2：无失效样本退化口径（MTBF 取运行小时，MTTR 取 0） —— //
    IF rFailCount < 0.5 THEN
        rMtbfH := rRunHours; // MTBF 取运行小时 [h] / MTBF equals running hours
        rMttrH := 0.0; // 无失效则无修复时间 / no failure, no repair time
        rAvailPct := rAvailCap; // 无失效窗内可用率按 100% 计 / availability capped at 100 percent
        iErrCode := 2; // 信息级：无失效样本 / info level: no failure sample
        bValid := TRUE;
        FC_DL_MtbfCalc := TRUE;
        RETURN;
    END_IF;
    rFailUse := rFailCount; // 生效失效次数 [次] / effective failure count
    // —— 段 3：量纲链 (h)/(次) = h —— //
    rMtbfRaw := rRunHours / rFailUse; // MTBF [h] / mean time between failures
    rMttrRaw := rRepairHours / rFailUse; // MTTR [h] / mean time to repair
    IF (ABS(rMtbfRaw) > 1.0E15) OR (ABS(rMttrRaw) > 1.0E15) THEN
        iErrCode := 3; // 结果非有限，强制归零 / non-finite result, forced to zero
        RETURN;
    END_IF;
    rMtbfH := rMtbfRaw;
    rMttrH := rMttrRaw;
    // —— 段 4：可用率（分母闸：MTBF+MTTR 不能为零） —— //
    rDenom := rMtbfH + rMttrH; // 分母 [h] / denominator
    IF ABS(rDenom) <= 1.0E-9 THEN
        rAvailPct := 0.0; // 分母退化，可用率置零 / degenerate denominator
        iErrCode := 3; // 信息级：可用率不可算 / info level: availability not computable
    ELSE
        rAvailPct := rMtbfH / rDenom * rInvPct; // 可用率 [%] / availability
        IF rAvailPct > rAvailCap THEN
            rAvailPct := rAvailCap; // 上限饱和 / saturate at cap
        ELSIF rAvailPct < 0.0 THEN
            rAvailPct := 0.0; // 下限钳零 / floor at zero
        END_IF
    END_IF;
    bValid := TRUE;
    FC_DL_MtbfCalc := TRUE;
END_FUNCTION

(* ---- FC_DL_OilChangeInterval.st ---- *)
(*
  道莅工业代码库 / Daoli Industrial ST Library
  组件: FC_DL_OilChangeInterval
  分类: DL_Device
  开源溯源: 无（clean-room 工程公式自研；参考公开工艺计算公式，未复制任何受版权保护代码）
  许可证: 本项目自有 (MIT)
  功能: 按负荷、温度、污染三因子修正换油周期，并给出剩余小时与到期判定
*)
FUNCTION FC_DL_OilChangeInterval : BOOL
VAR_INPUT
    rBaseHours : REAL; // 基准换油周期 [h] / base oil change interval
    rLoadFactor : REAL; // 负荷修正因子 [-]，域 (0.1, 5.0] / load correction factor
    rTempFactor : REAL; // 温度修正因子 [-]，域 (0.1, 5.0] / temperature correction factor
    rContamFactor : REAL; // 污染修正因子 [-]，域 (0.1, 5.0] / contamination correction factor
    rHoursSince : REAL; // 上次换油后已运行小时 [h] / hours since last oil change
END_VAR
VAR_OUTPUT
    rIntervalH : REAL; // 修正后换油周期 [h] / corrected interval
    rRemainH : REAL; // 剩余可用小时 [h]，可为负（已超期）/ remaining hours, negative when overdue
    bValid : BOOL; // 结果有效位 [-] / result valid flag
    bDue : BOOL; // 到期标志（剩余 ≤ 0）[-] / due flag
    iErrCode : INT; // 事件码 0=正常 1=修正因子超域 2=基准周期非法 3=结果非有限 / event code
END_VAR
VAR CONSTANT
    rFactorLo : REAL := 0.1; // 因子域下限（不含）[-] / factor domain lower bound, exclusive
    rFactorHi : REAL := 5.0; // 因子域上限（含）[-] / factor domain upper bound, inclusive
END_VAR
VAR
    rIntervalRaw : REAL; // 未校验周期 [h] / unchecked interval
END_VAR

    // —— 段 0：全路径预清 —— //
    rIntervalRaw := 0.0;
    rIntervalH := 0.0;
    rRemainH := 0.0;
    bValid := FALSE;
    bDue := FALSE;
    iErrCode := 0;
    FC_DL_OilChangeInterval := FALSE;
    // —— 段 1：三因子域闸（含非正因子，防周期符号翻转） —— //
    IF (rLoadFactor <= rFactorLo) OR (rLoadFactor > rFactorHi)
       OR (rTempFactor <= rFactorLo) OR (rTempFactor > rFactorHi)
       OR (rContamFactor <= rFactorLo) OR (rContamFactor > rFactorHi) THEN
        iErrCode := 1; // 修正因子超域，周期不可信 / correction factor out of domain
        RETURN;
    END_IF;
    // —— 段 2：基准周期域闸 —— //
    IF rBaseHours <= 0.0 THEN
        iErrCode := 2; // 基准周期非法，周期无定义 / invalid base interval
        RETURN;
    END_IF;
    // —— 段 3：量纲链 (h)×(-)×(-)×(-) = h —— //
    rIntervalRaw := rBaseHours * rLoadFactor * rTempFactor * rContamFactor; // 修正周期 [h] / corrected interval
    IF ABS(rIntervalRaw) > 1.0E15 THEN
        iErrCode := 3; // 结果非有限，强制归零 / non-finite result, forced to zero
        RETURN;
    END_IF;
    rIntervalH := rIntervalRaw;
    // —— 段 4：剩余小时（可为负，负值即超期量）与到期判定 —— //
    rRemainH := rIntervalH - rHoursSince; // 剩余小时 [h] / remaining hours
    bDue := rRemainH <= 0.0; // 到期判定 [-] / due test
    bValid := TRUE;
    FC_DL_OilChangeInterval := TRUE;
END_FUNCTION

(* ---- FC_DL_OrpRefOffsetCalc.st ---- *)
(* ============================================================
   DL_Device / FC_DL_OrpRefOffsetCalc ｜ v1.0.0 ｜ 2026-11-25
   功能：ORP 参比电位偏移修正 E_ref(T) = E_ref(25°C) + k·(T − 25) [mV]，
         fOffsetMv 为加到读数上换到 SHE 的修正量，fRefCorrMv = E_ref(T) − 实测参比。
   边界：nRefType ∉ {0,1,2} → 按 SHE（0 mV、k=0）处理并返回 FALSE；
         温度 ∉ [−5, 80]°C → 钳定并返回 FALSE（温补系数不外推）；
         任一浮点入参非有限 → 两出口同拍写 0（N1）。签名无出口码，故各闸
         一律以返回值 FALSE 上报，闸序即归因序（类型 → 非有限 → 温度）。
         量纲清单（N5）：k 单位 mV/°C；Ag/AgCl(3.5M KCl)=+0.20、饱和甘汞 SCE=+0.24、
         SHE=0.0；回代：25°C Ag/AgCl 标称 199 mV → E_SHE = E_meas + 199。
   依赖：仅 IEC 61131-3（无外部依赖，纯算术） ｜ 溯源：DLF-D-WATERANA
   验收：E_meas=550/T=25/标称 199/实测 199/类型 0 → 修正 199 mV、偏移 0 mV、TRUE；
         nRefType=7 → 按 SHE 折算（修正 0 mV）并返回 FALSE。
   ============================================================ *)
FUNCTION FC_DL_OrpRefOffsetCalc : BOOL
VAR_INPUT
    fMeasMv       : REAL;  // ORP 表实测读数（相对自身参比）[mV] / Measured ORP reading against its own reference
    fRefNominalMv : REAL;  // 参比标称电位（25°C 相对 SHE）[mV] / Nominal reference potential at twenty five Celsius
    fRefMeasMv    : REAL;  // 参比实测电位（相对 SHE）[mV] / Measured reference potential against the hydrogen electrode
    fSampleTempC  : REAL;  // 水样温度 [°C] / Sample temperature in Celsius degrees
    nRefType      : DINT;  // 参比类型 0=Ag/AgCl 1=SCE 2=SHE [-] / Reference electrode type selector
END_VAR
VAR_OUTPUT
    fOffsetMv  : REAL;  // 换算到 SHE 的修正量（加到读数上）[mV] / Correction added to the reading to reach SHE
    fRefCorrMv : REAL;  // 实测参比相对标称的偏移 [mV] / Measured reference deviation from the nominal value
END_VAR
VAR
    _fT    : REAL;  // 钳定后温度 [°C] / Clamped temperature
    _fK    : REAL;  // 温补系数 [mV/°C] / Temperature coefficient of the reference electrode
    _fNom  : REAL;  // 实际采用的参比标称电位 [mV] / Nominal reference potential actually used
    _fRefT : REAL;  // 温度修正后参比电位 [mV] / Temperature corrected reference potential
    _bTLim : BOOL;  // 温度越域标志 [-] / Temperature out of range flag
    _bType : BOOL;  // 参比类型非法标志 [-] / Illegal reference type flag
END_VAR
VAR CONSTANT
    DL_ORP_TREF   : REAL := 25.0;   // 参考温度 [°C] / Reference temperature
    DL_ORP_TLO    : REAL := -5.0;   // 温度域下限 [°C] / Lower temperature bound
    DL_ORP_THI    : REAL := 80.0;   // 温度域上限 [°C] / Upper temperature bound
    DL_ORP_K_AGCL : REAL := 0.20;   // Ag/AgCl 温补系数 [mV/°C] / Temperature coefficient of the silver chloride reference
    DL_ORP_K_SCE  : REAL := 0.24;   // 饱和甘汞温补系数 [mV/°C] / Temperature coefficient of the calomel reference
END_VAR

(* 段 0：出口预置安全侧（两出口 0，N1/N3） *)
FC_DL_OrpRefOffsetCalc := FALSE;
fOffsetMv := 0.0;  fRefCorrMv := 0.0;
_bTLim := FALSE;   _bType := FALSE;

(* 段 1：非有限闸（四个浮点入参；NaN 自反 + Inf 差值自减双判，R79/R272） *)
IF (fMeasMv <> fMeasMv) OR (fRefNominalMv <> fRefNominalMv)
   OR (fRefMeasMv <> fRefMeasMv) OR (fSampleTempC <> fSampleTempC) THEN RETURN; END_IF
IF ((fMeasMv - fMeasMv) <> (fMeasMv - fMeasMv))
   OR ((fRefNominalMv - fRefNominalMv) <> (fRefNominalMv - fRefNominalMv))
   OR ((fRefMeasMv - fRefMeasMv) <> (fRefMeasMv - fRefMeasMv))
   OR ((fSampleTempC - fSampleTempC) <> (fSampleTempC - fSampleTempC)) THEN RETURN; END_IF

(* 段 2：参比类型分派（非法按 SHE，k=0、基准 0 mV） *)
CASE nRefType OF
0:      _fK := DL_ORP_K_AGCL;  _fNom := fRefNominalMv;
1:      _fK := DL_ORP_K_SCE;   _fNom := fRefNominalMv;
2:      _fK := 0.0;            _fNom := 0.0;
ELSE
    _fK := 0.0;  _fNom := 0.0;  _bType := TRUE;   // 非法类型：按 SHE 折算
END_CASE

(* 段 3：温度域闸（越域钳定，禁外推） *)
_fT := fSampleTempC;
IF fSampleTempC < DL_ORP_TLO THEN
    _fT := DL_ORP_TLO;  _bTLim := TRUE;
ELSIF fSampleTempC > DL_ORP_THI THEN
    _fT := DL_ORP_THI;  _bTLim := TRUE;
END_IF

(* 段 4：温度修正后的参比电位与偏移（乘加，无除法） *)
_fRefT := _fNom + _fK * (_fT - DL_ORP_TREF);

(* 段 5：单一出口裁决（两出口同源赋值一次，N4） *)
fOffsetMv  := _fRefT;
fRefCorrMv := _fRefT - fRefMeasMv;
IF (fOffsetMv <> fOffsetMv) OR (fRefCorrMv <> fRefCorrMv)
   OR ((fOffsetMv - fOffsetMv) <> (fOffsetMv - fOffsetMv))
   OR ((fRefCorrMv - fRefCorrMv) <> (fRefCorrMv - fRefCorrMv)) THEN
    fOffsetMv := 0.0;  fRefCorrMv := 0.0;   // 出口非有限：实值同拍写 0 且返回 FALSE（N1）
    RETURN;
END_IF
IF _bType OR _bTLim THEN
    FC_DL_OrpRefOffsetCalc := FALSE;    // 类型非法/温度越域：值照给，供上层记录
    RETURN;
END_IF
FC_DL_OrpRefOffsetCalc := TRUE;
END_FUNCTION

(* ---- FC_DL_PadWearIndexCalc.st ---- *)
(*
  ============================================================
  组件名 : FC_DL_PadWearIndexCalc
  分类   : DL_Device
  功能   : 吸盘磨损指数计算，综合泄漏增长率与直径磨耗量加权后给出更换到期判定
  复杂度 : C2
  版本   : 1.0.0
  作者   : 道莅工业代码库工厂 / R81
  日期   : 2026-11-24
  开源溯源 : clean-room（no upstream）—— 依据公开工程公式自研，未复制任何上游实现
  红线自检 : R1 无GVL/R2 无物理地址/R3 纯IEC/R4 防除零/R5 双语注释
  接口说明 :
      泄漏增长率 = (当前泄漏 - 新品泄漏) / 新品泄漏 * 100，新品泄漏低于 0.001 L/min 视为无基准判无效。
      磨损指数 = 0.7 * 泄漏增长率 + 0.3 * 直径磨耗 * 10，限幅 0~100。
      指数超过 70 判更换到期；负的泄漏增长（密封变好）按 0 截断，指数只反映劣化方向。
  ============================================================
*)
FUNCTION FC_DL_PadWearIndexCalc : BOOL
VAR_INPUT
    bEnable     : BOOL; // 使能：TRUE 时计算 / Enable: TRUE to compute
    bErr        : BOOL; // 外部故障：TRUE 时立即退出并置结果无效 / External fault: TRUE aborts with invalid result
    rLeakNew    : REAL; // 新品基准泄漏量 [L/min] / leak rate of a new pad [litre per minute]
    rLeakNow    : REAL; // 当前实测泄漏量 [L/min] / currently measured leak rate [litre per minute]
    rDiaWear_mm : REAL; // 吸盘直径磨耗量 [mm] / diameter wear of the pad [millimetre]
END_VAR
VAR_OUTPUT
    rLeakPct  : REAL; // 泄漏增长率 [%] / leak growth rate [percent]
    rWearIdx  : REAL; // 综合磨损指数，限幅 0~100 [无量纲] / combined wear index clamped to 0 to 100 [dimensionless]
    bReplaceDue : BOOL; // 更换到期：TRUE 表示指数超过 70 / replacement due, TRUE when the index exceeds 70
    bValid    : BOOL; // 输出有效：TRUE 表示结果可用 / Output valid
END_VAR
VAR CONSTANT
    DL_R_MAX     : REAL := 3.0E38;  // 实数上界，用于拦截 Inf [无量纲] / real upper bound used to reject infinity [dimensionless]
    DL_EPS       : REAL := 1.0E-12; // 除零判定阈值 [无量纲] / division guard threshold [dimensionless]
    DL_LEAK_MIN  : REAL := 0.001;   // 新品泄漏基准的可信下界 [L/min] / credible lower bound of the new pad leak reference [litre per minute]
    DL_PCT       : REAL := 100.0;   // 百分数换算系数 [无量纲] / percentage scaling factor [dimensionless]
    DL_W_LEAK    : REAL := 0.7;     // 泄漏项权重 [无量纲] / weight of the leak term [dimensionless]
    DL_W_DIA     : REAL := 0.3;     // 直径磨耗项权重 [无量纲] / weight of the diameter wear term [dimensionless]
    DL_DIA_GAIN  : REAL := 10.0;    // 直径磨耗放大倍数 [无量纲] / amplification of the diameter wear term [dimensionless]
    DL_IDX_HI    : REAL := 100.0;   // 指数限幅上限 [无量纲] / upper clamp of the index [dimensionless]
    DL_IDX_LO    : REAL := 0.0;     // 指数限幅下限 [无量纲] / lower clamp of the index [dimensionless]
    DL_DUE_IDX   : REAL := 70.0;    // 更换到期门限 [无量纲] / replacement due threshold [dimensionless]
    DL_DIA_MAX   : REAL := 200.0;   // 直径磨耗合理上限 [mm] / sanity upper bound of the diameter wear [millimetre]
END_VAR
VAR
    _bFin : BOOL := FALSE; // 输入有限性判定结果 / input finiteness verdict
    _rRaw : REAL := 0.0;   // 限幅前磨损指数 [无量纲] / raw wear index before clamping [dimensionless]
END_VAR

    // 段 1｜出口预置
    rLeakPct := 0.0;
    rWearIdx := 0.0;
    bReplaceDue := FALSE;
    bValid := FALSE;
    // 段 2｜使能闸与外部故障闸
    IF NOT bEnable THEN
        RETURN;
    END_IF;
    IF bErr THEN
        RETURN;
    END_IF;
    // 段 3｜非有限闸
    _bFin := (rLeakNew = rLeakNew) AND (ABS(rLeakNew) <= DL_R_MAX) AND (rLeakNow = rLeakNow) AND (ABS(rLeakNow) <= DL_R_MAX) AND (rDiaWear_mm = rDiaWear_mm) AND (ABS(rDiaWear_mm) <= DL_R_MAX);
    IF NOT _bFin THEN
        RETURN;
    END_IF;
    // 段 4｜域闸：新品泄漏必须高于可信下界，当前泄漏与磨耗不得为负
    IF (ABS(rLeakNew) <= DL_EPS) OR (rLeakNew < DL_LEAK_MIN) THEN
        RETURN;
    END_IF;
    IF (rLeakNow < 0.0) OR (rDiaWear_mm < 0.0) OR (rDiaWear_mm > DL_DIA_MAX) THEN
        RETURN;
    END_IF;
    // 段 5｜泄漏增长率
    rLeakPct := (rLeakNow - rLeakNew) / rLeakNew * DL_PCT;
    IF rLeakPct < DL_IDX_LO THEN
        rLeakPct := DL_IDX_LO;
    END_IF;
    // 段 6｜加权合成与限幅
    _rRaw := DL_W_LEAK * rLeakPct + DL_W_DIA * rDiaWear_mm * DL_DIA_GAIN;
    IF _rRaw < DL_IDX_LO THEN
        rWearIdx := DL_IDX_LO;
    ELSIF _rRaw > DL_IDX_HI THEN
        rWearIdx := DL_IDX_HI;
    ELSE
        rWearIdx := _rRaw;
    END_IF;
    // 段 7｜更换到期判定用限幅前的真实指数判断方向
    IF _rRaw > DL_DUE_IDX THEN
        bReplaceDue := TRUE;
    ELSE
        bReplaceDue := FALSE;
    END_IF;
    bValid := TRUE;
    FC_DL_PadWearIndexCalc := bValid;
END_FUNCTION

(* ---- FC_DL_PaintConsumptionCalc.st ---- *)
(*
  Name: FC_DL_PaintConsumptionCalc
  Category: DL_Device
  Version: 1.0.0
  Round: R89 / 2026-11-25
  开源溯源：clean-room 自研（族 涂装喷涂线，ST 开源生态实测 0 命中，无外部代码引入）
  功能：单件涂料消耗与利用率：实际用量按流量×节拍÷件数折算，理论用量按膜厚×面积÷固含量折算。
  边界条件：① 六入参全部过非有限闸，任一非有限返回哨兵 -1；
            ② 件数为除子（≥ 1 件）、固含量为除子（5~100 %）、面积为理论用量乘数，全部域闸拦截；
            ③ 利用率 = 理论湿漆量 ÷ 实际用量 × 100，可超 100 %（表明实际用量偏低，照实上报不钳位）。
  量纲自证：ml/min × s ÷ 60 = ml；μm × m2 = ml（1 μm·m2 = 1 ml）；两者同量纲故比值无量纲。
*)
FUNCTION FC_DL_PaintConsumptionCalc : REAL
VAR_INPUT
    fFlowMlmin : REAL;      (* 喷枪湿漆流量 [ml/min] Wet paint flow [ml/min] *)
    fCycleTimeS : REAL;     (* 单次喷涂节拍 [s] Coating cycle time [s] *)
    nParts : INT;           (* 单次节拍内件数 [件] Parts per cycle *)
    fSolidPct : REAL;       (* 固含量（质量） [%] Solids content [%] *)
    fFilmUm : REAL;         (* 目标干膜厚度 [μm] Target dry film thickness [um] *)
    fAreaM2 : REAL;         (* 单件喷涂面积 [m2] Coated area per part [m2] *)
END_VAR
VAR_OUTPUT
    fPaintPerPartMl : REAL; (* 单件实际消耗 [ml] Paint consumption per part [ml] *)
    fUtilPct : REAL;        (* 涂料利用率 [%] Paint utilization [%] *)
    xValid : BOOL;          (* 计算有效性标志 [-] Calculation valid flag *)
END_VAR
VAR CONSTANT
    DL_EPS : REAL := 1.0E-9;        (* 判据容差 [-] Criterion tolerance *)
    DL_SECMIN : REAL := 60.0;       (* 每秒 → 每分钟换算 [s/min] Second to minute *)
    DL_PCT : REAL := 100.0;         (* 百分数基准 [%] Percent base *)
    DL_F_MIN : REAL := 1.0;         (* 流量下限 [ml/min] Flow floor [ml/min] *)
    DL_F_MAX : REAL := 2000.0;      (* 流量上限 [ml/min] Flow ceiling [ml/min] *)
    DL_T_MIN : REAL := 1.0;         (* 节拍下限 [s] Cycle floor [s] *)
    DL_T_MAX : REAL := 3600.0;      (* 节拍上限 [s] Cycle ceiling [s] *)
    DL_N_MAX : INT := 500;          (* 件数上限 [件] Part count ceiling *)
    DL_S_MIN : REAL := 5.0;         (* 固含量下限 [%] Solids floor [%] *)
    DL_S_MAX : REAL := 100.0;       (* 固含量上限 [%] Solids ceiling [%] *)
    DL_FILM_MIN : REAL := 1.0;      (* 膜厚下限 [μm] Film floor [um] *)
    DL_FILM_MAX : REAL := 200.0;    (* 膜厚上限 [μm] Film ceiling [um] *)
    DL_A_MIN : REAL := 0.001;       (* 面积下限 [m2] Area floor [m2] *)
    DL_A_MAX : REAL := 100.0;       (* 面积上限 [m2] Area ceiling [m2] *)
END_VAR
VAR
    fActualMl : REAL;   (* 单次节拍实际用量 [ml] Actual paint per cycle [ml] *)
    fTheoryMl : REAL;   (* 单件理论湿漆量 [ml] Theoretical wet paint per part [ml] *)
END_VAR
(* 出口预置：三出口统一预置（R256） *)
fPaintPerPartMl := 0.0; fUtilPct := 0.0; xValid := FALSE;
(* 非有限闸：NaN 自反判 + Inf 差值自减判，五浮点入参全枚举（R272） *)
IF (fFlowMlmin <> fFlowMlmin) OR ((fFlowMlmin - fFlowMlmin) <> 0.0)
   OR (fCycleTimeS <> fCycleTimeS) OR ((fCycleTimeS - fCycleTimeS) <> 0.0)
   OR (fSolidPct <> fSolidPct) OR ((fSolidPct - fSolidPct) <> 0.0)
   OR (fFilmUm <> fFilmUm) OR ((fFilmUm - fFilmUm) <> 0.0)
   OR (fAreaM2 <> fAreaM2) OR ((fAreaM2 - fAreaM2) <> 0.0) THEN
    FC_DL_PaintConsumptionCalc := -1.0;     (* 哨兵 -1：入参非有限 / Sentinel -1, non-finite input *)
    RETURN;
END_IF
(* 组态域闸：流量、节拍、件数、固含量、膜厚、面积逐项定域（件数与固含为除子） *)
IF (fFlowMlmin < DL_F_MIN) OR (fFlowMlmin > DL_F_MAX)
   OR (fCycleTimeS < DL_T_MIN) OR (fCycleTimeS > DL_T_MAX)
   OR (nParts < 1) OR (nParts > DL_N_MAX)
   OR (fSolidPct < DL_S_MIN) OR (fSolidPct > DL_S_MAX)
   OR (fFilmUm < DL_FILM_MIN) OR (fFilmUm > DL_FILM_MAX)
   OR (fAreaM2 < DL_A_MIN) OR (fAreaM2 > DL_A_MAX) THEN
    FC_DL_PaintConsumptionCalc := -1.0;     (* 哨兵 -1：组态非法 / Sentinel -1, bad configuration *)
    RETURN;
END_IF
(* 单次节拍实际用量：ml/min × s ÷ 60 = ml *)
fActualMl := fFlowMlmin * fCycleTimeS / DL_SECMIN;
(* 单件实际用量：件数已过下限闸，绝无零除 *)
fPaintPerPartMl := fActualMl / INT_TO_REAL(nParts);
(* 单件理论湿漆量：膜厚[μm] × 面积[m2] = ml（湿体积），再除固含量折算湿漆 *)
fTheoryMl := (fFilmUm * fAreaM2) / (fSolidPct / DL_PCT);
(* 利用率：理论 ÷ 实际 × 100，实际用量已由流量下限保证为正 *)
fUtilPct := (fTheoryMl / fPaintPerPartMl) * DL_PCT;
xValid := TRUE;                             (* 链路有效 / Chain valid *)
FC_DL_PaintConsumptionCalc := fPaintPerPartMl;
END_FUNCTION

(* ---- FC_DL_PaintFilmThicknessCalc.st ---- *)
(*
  Name: FC_DL_PaintFilmThicknessCalc
  Category: DL_Device
  Version: 1.0.0
  Round: R89 / 2026-11-25
  开源溯源：clean-room 自研（族 涂装喷涂线，ST 开源生态实测 0 命中，无外部代码引入）
  功能：漆膜厚度估算：湿漆流量 × 密度 × 固含量 ÷ 干膜密度 ÷ 单位时间喷涂面积 = 干膜厚度。
  边界条件：① 四入参全部过非有限闸，任一非有限返回哨兵 -1；
            ② 喷涂面积为除子，按 0.01~100 m2/min 域闸拦截，绝无零除；
            ③ 干膜密度取常量 DL_PFT_RHO_FILM = 1.2 g/cm3（通用涂料干膜密度），属工艺常量非实测；
            ④ 固含量按下限 5 % 域闸拦截，避免固含趋零导致膜厚趋零的伪结论。
  量纲自证：ml/min × g/ml = g/min；× 固含 = 固体 g/min；÷ g/cm3 = cm3/min；÷ m2/min = cm3/m2，
            而 1 cm3 均布于 1 m2 即 1 μm，故数值直接为 μm。
*)
FUNCTION FC_DL_PaintFilmThicknessCalc : REAL
VAR_INPUT
    fFlowMlmin : REAL;          (* 湿漆流量 [ml/min] Wet paint flow [ml/min] *)
    fSolidPct : REAL;           (* 固含量（质量） [%] Solids content by mass [%] *)
    fAreaM2min : REAL;          (* 单位时间喷涂面积 [m2/min] Coated area per minute [m2/min] *)
    fDensityGml : REAL;         (* 湿漆密度 [g/ml] Wet paint density [g/ml] *)
END_VAR
VAR_OUTPUT
    fFilmUm : REAL;             (* 干膜厚度 [μm] Dry film thickness [um] *)
    xValid : BOOL;              (* 计算有效性标志 [-] Calculation valid flag *)
END_VAR
VAR CONSTANT
    DL_EPS : REAL := 1.0E-9;        (* 判据容差 [-] Criterion tolerance *)
    DL_PFT_RHO_FILM : REAL := 1.2;  (* 干膜密度（工艺常量） [g/cm3] Dry film density [g/cm3] *)
    DL_PCT : REAL := 100.0;         (* 百分数基准 [%] Percent base *)
    DL_F_MIN : REAL := 1.0;         (* 流量下限 [ml/min] Flow floor [ml/min] *)
    DL_F_MAX : REAL := 2000.0;      (* 流量上限 [ml/min] Flow ceiling [ml/min] *)
    DL_S_MIN : REAL := 5.0;         (* 固含量下限 [%] Solids floor [%] *)
    DL_S_MAX : REAL := 100.0;       (* 固含量上限 [%] Solids ceiling [%] *)
    DL_A_MIN : REAL := 0.01;        (* 面积下限 [m2/min] Area floor [m2/min] *)
    DL_A_MAX : REAL := 100.0;       (* 面积上限 [m2/min] Area ceiling [m2/min] *)
    DL_D_MIN : REAL := 0.7;         (* 湿漆密度下限 [g/ml] Density floor [g/ml] *)
    DL_D_MAX : REAL := 2.0;         (* 湿漆密度上限 [g/ml] Density ceiling [g/ml] *)
END_VAR
VAR
    fSolidGmin : REAL;  (* 固体质量流量 [g/min] Solids mass flow [g/min] *)
    fVolCm3min : REAL;  (* 固体体积流量 [cm3/min] Solids volume flow [cm3/min] *)
END_VAR
(* 出口预置：两出口统一预置（R256） *)
fFilmUm := 0.0; xValid := FALSE;
(* 非有限闸：NaN 自反判 + Inf 差值自减判，四入参全枚举 *)
IF (fFlowMlmin <> fFlowMlmin) OR ((fFlowMlmin - fFlowMlmin) <> 0.0)
   OR (fSolidPct <> fSolidPct) OR ((fSolidPct - fSolidPct) <> 0.0)
   OR (fAreaM2min <> fAreaM2min) OR ((fAreaM2min - fAreaM2min) <> 0.0)
   OR (fDensityGml <> fDensityGml) OR ((fDensityGml - fDensityGml) <> 0.0) THEN
    FC_DL_PaintFilmThicknessCalc := -1.0;   (* 哨兵 -1：入参非有限 / Sentinel -1, non-finite input *)
    RETURN;
END_IF
(* 组态域闸：流量、固含量、面积为除子、密度逐项定域 *)
IF (fFlowMlmin < DL_F_MIN) OR (fFlowMlmin > DL_F_MAX)
   OR (fSolidPct < DL_S_MIN) OR (fSolidPct > DL_S_MAX)
   OR (fAreaM2min < DL_A_MIN) OR (fAreaM2min > DL_A_MAX)
   OR (fDensityGml < DL_D_MIN) OR (fDensityGml > DL_D_MAX) THEN
    FC_DL_PaintFilmThicknessCalc := -1.0;   (* 哨兵 -1：组态非法 / Sentinel -1, bad configuration *)
    RETURN;
END_IF
(* 固体质量流量：ml/min × g/ml = g/min，再乘固含比例 *)
fSolidGmin := fFlowMlmin * fDensityGml * (fSolidPct / DL_PCT);
(* 固体体积流量：g/min ÷ g/cm3 = cm3/min，干膜密度为常量恒正 *)
fVolCm3min := fSolidGmin / DL_PFT_RHO_FILM;
(* 膜厚：cm3/min ÷ m2/min = cm3/m2 ≡ μm，面积已过下限闸 *)
fFilmUm := fVolCm3min / fAreaM2min;
xValid := TRUE;                             (* 链路有效 / Chain valid *)
FC_DL_PaintFilmThicknessCalc := fFilmUm;
END_FUNCTION

(* ---- FC_DL_PalletOverhangCalc.st ---- *)
(*
  DL Factory R83 | FC_DL_PalletOverhangCalc
  功能：算托盘相对货垛的单侧悬垂量，并按允许悬垂比例校验堆码稳定性。
  开源溯源：无（clean-room 自研，依据公开工艺公式，来源=行业通用公式，许可证=MIT，借鉴点=公式结构）
  规则：R1-R21 全遵守
*)
FUNCTION FC_DL_PalletOverhangCalc : REAL
VAR_INPUT
    fPalletLenMm : REAL; // 托盘长度 [mm] / Pallet length [mm]
    fPalletWidMm : REAL; // 托盘宽度 [mm] / Pallet width [mm]
    fBoxLenMm    : REAL; // 货垛沿长度方向外形尺寸 [mm] / Load footprint length [mm]
    fBoxWidMm    : REAL; // 货垛沿宽度方向外形尺寸 [mm] / Load footprint width [mm]
    fMaxOverPct  : REAL; // 允许单侧悬垂比例（0~10）[%] / Allowed overhang ratio [%]
END_VAR
VAR_OUTPUT
    fOverLenMm : REAL; // 长度方向单侧悬垂（负值=货垛内缩）[mm] / Length overhang [mm]
    fOverWidMm : REAL; // 宽度方向单侧悬垂 [mm] / Width overhang [mm]
    fOverMaxMm : REAL; // 该托盘允许的单侧悬垂上限（两向较严者）[mm] / Allowed ceiling [mm]
    xOk        : BOOL; // 悬垂合规判定 / Overhang compliance flag
    xValid     : BOOL; // 计算有效性标志 / Calculation validity flag
END_VAR
VAR
    fLimLenMm : REAL; // 长度向允许悬垂 [mm] / Allowed overhang on length [mm]
    fLimWidMm : REAL; // 宽度向允许悬垂 [mm] / Allowed overhang on width [mm]
END_VAR
fOverLenMm := 0.0; fOverWidMm := 0.0; fOverMaxMm := 0.0; xOk := FALSE; xValid := FALSE; // 出口预置
// 非有限拦截 + 量纲自检（R20/R21）
IF NOT (fPalletLenMm > -1.0E30 AND fPalletLenMm < 1.0E30) OR NOT (fPalletWidMm > -1.0E30 AND fPalletWidMm < 1.0E30) OR NOT (fBoxLenMm > -1.0E30 AND fBoxLenMm < 1.0E30) OR NOT (fBoxWidMm > -1.0E30 AND fBoxWidMm < 1.0E30) OR NOT (fMaxOverPct > -1.0E30 AND fMaxOverPct < 1.0E30) OR fPalletLenMm <= 0.0 OR fPalletWidMm <= 0.0 OR fBoxLenMm <= 0.0 OR fBoxWidMm <= 0.0 OR fMaxOverPct < 0.0 THEN
    FC_DL_PalletOverhangCalc := -1.0; RETURN;  // 哨兵 -1：非有限或量纲越界 / Sentinel -1
END_IF
// 悬垂比例域闸：0~10% 之外钳位（超 10% 已无稳定可言）
IF fMaxOverPct > 10.0 THEN
    fMaxOverPct := 10.0;            // 上限钳位 [%] / Clamp upper bound
END_IF
// 单侧悬垂：两向外形差 ÷ 2，同量纲（mm）相减；负值表示货垛内缩
fOverLenMm := (fPalletLenMm - fBoxLenMm) / 2.0;   // 长度向单侧悬垂 [mm] / Length overhang [mm]
fOverWidMm := (fPalletWidMm - fBoxWidMm) / 2.0;   // 宽度向单侧悬垂 [mm] / Width overhang [mm]
// 允许上限：托盘该向尺寸 × 比例 ÷ 100（mm × 无量纲 = mm，量纲自洽）
fLimLenMm := fPalletLenMm * (fMaxOverPct / 100.0); // 长度向允许悬垂 [mm] / Allowed length overhang
fLimWidMm := fPalletWidMm * (fMaxOverPct / 100.0); // 宽度向允许悬垂 [mm] / Allowed width overhang
// 上限回显取两向较严者，供上层 HMI 统一显示
IF fLimLenMm <= fLimWidMm THEN
    fOverMaxMm := fLimLenMm;        // 长度向更严 [mm] / Length direction is stricter
ELSE
    fOverMaxMm := fLimWidMm;        // 宽度向更严 [mm] / Width direction is stricter
END_IF
// 合规判定：两向悬垂均不超各自上限（负值内缩恒合规）
xOk    := (fOverLenMm <= fLimLenMm) AND (fOverWidMm <= fLimWidMm); // 合规布尔 / Compliance boolean
xValid := TRUE; FC_DL_PalletOverhangCalc := fOverLenMm; // 返回长度向悬垂 [mm] / Return overhang
END_FUNCTION

(* ---- FC_DL_PhAsymmPotentialCalc.st ---- *)
(* ============================================================
   DL_Device / FC_DL_PhAsymmPotentialCalc ｜ v1.0.0 ｜ 2026-11-25
   功能：pH 零点不对称电位 E_asym = mV_meas + S(T)·(pH − 7.00) [mV]，
         S(T) = 59.16 × (273.15 + T) / 298.15 [mV/pH]（Nernst 温度修正）。
   边界：温度 ∉ [−5, 80]°C → 钳定后计算并报码 1（温补系数不许外推）；
         任一入参非有限 → 码 2、出口写 0（N1：判据与实值同源落安全侧）；
         |E_asym| > 30 mV → 码 3（电极钝化/污染），值照给供上层告警。
   依赖：仅 IEC 61131-3（ABS） ｜ 溯源：DLF-D-WATERANA（内部原创线）
   验收：mV=3.0/pH=7.00/T=25 → +3.0 mV、码 0；mV=+62.16/pH=6.00/T=25 →
         62.16 − 59.16 = +3.0 mV；T=100 → 钳到 80°C 计算、码 1（不外推）。
   ============================================================ *)
FUNCTION FC_DL_PhAsymmPotentialCalc : BOOL
VAR_INPUT
    fMvMeas : REAL;  // 电极实测电位 [mV] / Measured electrode potential in millivolts
    fPhMeas : REAL;  // 实测 pH 值（同点采样）[pH] / Measured pH value taken at the same instant
    fTempC  : REAL;  // 溶液温度 [°C] / Solution temperature in Celsius degrees
END_VAR
VAR_OUTPUT
    fAsymmV : REAL;   // 不对称电位（零点偏移）[mV] / Asymmetry potential, the zero point shift
    uErrId  : UDINT;  // 码 0 正常 / 1 温度越域 / 2 非有限 / 3 不对称超 30 mV [-] / Outlet code
END_VAR
VAR
    _fT     : REAL;  // 钳定后温度 [°C] / Clamped temperature
    _fSlope : REAL;  // 温度修正后理论斜率 [mV/pH] / Temperature corrected theoretical slope
    _fAsym  : REAL;  // 不对称电位中间值 [mV] / Intermediate asymmetry potential
    _bTLim  : BOOL;  // 温度越域标志 [-] / Temperature out of range flag
END_VAR
VAR CONSTANT
    DL_PHA_S25   : REAL := 59.16;   // 25 摄氏度理论斜率 [mV/pH] / Theoretical slope at twenty five Celsius
    DL_PHA_TREF  : REAL := 25.0;    // 参考温度 [°C] / Reference temperature
    DL_PHA_TK    : REAL := 273.15;  // 绝对零度偏移 [K] / Kelvin offset of the Celsius scale
    DL_PHA_TPT7  : REAL := 7.00;    // pH 零点 [pH] / Neutral pH reference point
    DL_PHA_TLO   : REAL := -5.0;    // 温度域下限 [°C] / Lower temperature bound
    DL_PHA_THI   : REAL := 80.0;    // 温度域上限 [°C] / Upper temperature bound
    DL_PHA_AMAX  : REAL := 30.0;    // 不对称电位接收上限 [mV] / Acceptance bound of the asymmetry
END_VAR

(* 段 0：出口预置安全侧（0 mV、码取最严，N1/N3） *)
FC_DL_PhAsymmPotentialCalc := FALSE;
fAsymmV := 0.0;  uErrId := 2;  _bTLim := FALSE;

(* 段 1：非有限闸（三入参 + 温度差） *)
IF (fMvMeas <> fMvMeas) OR (fPhMeas <> fPhMeas) OR (fTempC <> fTempC) THEN RETURN; END_IF
IF ((fTempC - fTempC) <> (fTempC - fTempC)) THEN RETURN; END_IF

(* 段 2：温度域闸（越域钳定并报码，禁外推） *)
_fT := fTempC;
IF fTempC < DL_PHA_TLO THEN
    _fT := DL_PHA_TLO;  _bTLim := TRUE;
ELSIF fTempC > DL_PHA_THI THEN
    _fT := DL_PHA_THI;  _bTLim := TRUE;
END_IF

(* 段 3：斜率与不对称电位（除子 298.15 为常量非零） *)
_fSlope := DL_PHA_S25 * (_fT + DL_PHA_TK) / (DL_PHA_TREF + DL_PHA_TK);
_fAsym  := fMvMeas + _fSlope * (fPhMeas - DL_PHA_TPT7);

(* 段 4：结果复检（非有限保持段 0 安全侧） *)
IF (_fAsym <> _fAsym) OR ((_fAsym - _fAsym) <> (_fAsym - _fAsym)) THEN RETURN; END_IF

(* 段 5：单一出口裁决（判据与出口同源于 _fAsym，N4/R23） *)
fAsymmV := _fAsym;
IF _bTLim THEN
    uErrId := 1;                        // 温度越域：值照给（已钳），FALSE 供上层记录
ELSIF ABS(_fAsym) > DL_PHA_AMAX THEN
    uErrId := 3;                        // 电极失效判据：值照给供上层告警
ELSE
    uErrId := 0;  FC_DL_PhAsymmPotentialCalc := TRUE;
END_IF
END_FUNCTION

(* ---- FC_DL_PhSlopeEffCalc.st ---- *)
(* ============================================================
   DL_Device / FC_DL_PhSlopeEffCalc ｜ v1.0.0 ｜ 2026-11-25
   功能：pH 电极斜率效率 fSlopePct = |S| / 59.16 × 100 [%]，
         S = (mV2 − mV1) / (pH2 − pH1) [mV/pH]，正常电极 S 为负值。
   边界：|ΔpH| ≤ 0.01 → 码 1（效率 0）；任一入参非有限 → 码 2（效率 0，N1 同拍改写）；
         效率 ∉ [85, 115]% → 码 3（效率照给 + bOutOfLim）。理论斜率取 25°C 名义
         59.16 mV/pH（R95 代理假设：覆盖 15~35°C 常规水样；恒温高精度场合由
         调用方按 Nernst 式补正后回灌，本件签名无温度引脚，不做温度修正）。
   依赖：仅 IEC 61131-3（ABS） ｜ 溯源：DLF-D-WATERANA（内部原创线）
   验收：mV1=0/pH1=7.00、mV2=+177.5/pH2=4.00 → S=−59.17、效率 100.0%、码 0；
         pH1=pH2 → 码 1、效率 0；效率 120% → 码 3、bOutOfLim=TRUE。
   ============================================================ *)
FUNCTION FC_DL_PhSlopeEffCalc : BOOL
VAR_INPUT
    fMv1 : REAL;  // 标定点 1 电极电位 [mV] / Electrode potential of calibration point one
    fPh1 : REAL;  // 标定点 1 的 pH 值 [pH] / pH value of calibration point one
    fMv2 : REAL;  // 标定点 2 电极电位 [mV] / Electrode potential of calibration point two
    fPh2 : REAL;  // 标定点 2 的 pH 值 [pH] / pH value of calibration point two
END_VAR
VAR_OUTPUT
    fSlopePct : REAL;   // 斜率效率 [%] / Slope efficiency in percent
    uErrId    : UDINT;  // 码 0 正常 / 1 两点重合 / 2 非有限 / 3 效率越限 [-] / Outlet code
    bOutOfLim : BOOL;   // 效率越出 85~115% [-] / Efficiency outside the acceptance band
END_VAR
VAR
    _fDph : REAL;  // pH 差 pH2 − pH1 [pH] / pH difference of the two points
    _fS   : REAL;  // 实测斜率 [mV/pH] / Measured slope in millivolts per pH
    _fEff : REAL;  // 效率中间值 [%] / Intermediate efficiency value
END_VAR
VAR CONSTANT
    DL_PHS_THEORY : REAL := 59.16;  // 25 摄氏度理论斜率 [mV/pH] / Theoretical slope at twenty five Celsius
    DL_PHS_MIND   : REAL := 0.01;   // 两点最小 pH 差 [pH] / Minimum pH distance of the two points
    DL_PHS_LO     : REAL := 85.0;   // 效率接收下限 [%] / Lower acceptance bound
    DL_PHS_HI     : REAL := 115.0;  // 效率接收上限 [%] / Upper acceptance bound
    DL_PHS_HUND   : REAL := 100.0;  // 百分比换算系数 [%] / Percent conversion factor
END_VAR

(* 段 0：出口预置安全侧（效率 0、越限置位，N1/N3） *)
FC_DL_PhSlopeEffCalc := FALSE;
fSlopePct := 0.0;  uErrId := 2;  bOutOfLim := TRUE;

(* 段 1：非有限闸（四入参 + 电位差） *)
IF (fMv1 <> fMv1) OR (fPh1 <> fPh1) OR (fMv2 <> fMv2) OR (fPh2 <> fPh2) THEN RETURN; END_IF
IF ((fMv2 - fMv1) - (fMv2 - fMv1)) <> ((fMv2 - fMv1) - (fMv2 - fMv1)) THEN RETURN; END_IF

(* 段 2：两点可分辨（pH 差域闸，防除零） *)
_fDph := fPh2 - fPh1;
IF ABS(_fDph) <= DL_PHS_MIND THEN uErrId := 1; RETURN; END_IF

(* 段 3：斜率与效率（除子已证 |ΔpH| > 0.01） *)
_fS   := (fMv2 - fMv1) / _fDph;
_fEff := ABS(_fS) / DL_PHS_THEORY * DL_PHS_HUND;
IF (_fEff <> _fEff) OR ((_fEff - _fEff) <> (_fEff - _fEff)) THEN RETURN; END_IF

(* 段 4：单一出口裁决（判据与出口同源于 _fEff，N4/R23） *)
fSlopePct := _fEff;
bOutOfLim := ((_fEff < DL_PHS_LO) OR (_fEff > DL_PHS_HI));
IF bOutOfLim THEN
    uErrId := 3;                        // 越限：效率照给，返回值 FALSE 供上层告警
ELSE
    uErrId := 0;  FC_DL_PhSlopeEffCalc := TRUE;
END_IF
END_FUNCTION

(* ---- FC_DL_PmScheduleNext.st ---- *)
(*
  道莅工业代码库 / Daoli Industrial ST Library
  组件: FC_DL_PmScheduleNext
  分类: DL_Device
  开源溯源: 无（clean-room 工程公式自研；参考公开工艺计算公式，未复制任何受版权保护代码）
  许可证: 本项目自有 (MIT)
  功能: 由上次 PM 时刻与周期天数推算下次 PM 时刻、下次 PM 日期与逾期天数
  时基声明: 时刻统一经 DT_TO_DINT 折算为「自 1970-01-01 起的秒计数」做整数运算，
            避免 TIME 型毫秒量在 24.8 天以上溢出 DINT；最大 3650 d × 86400 s = 3.15E8 s 安全
*)
FUNCTION FC_DL_PmScheduleNext : BOOL
VAR_INPUT
    dtLast : DT; // 上次 PM 完成时刻 [DT] / last PM completion timestamp
    dtNow : DT; // 当前时刻 [DT] / current timestamp
    iIntervalDays : INT; // PM 周期 [d]，域 (0, 3650] / PM interval in days
END_VAR
VAR_OUTPUT
    dtNext : DT; // 下次 PM 到期时刻 [DT] / next PM due timestamp
    dNextDate : DATE; // 下次 PM 到期日期 [DATE] / next PM due date, operator friendly
    iOverdueDays : INT; // 逾期天数 [d]，未逾期为 0 / overdue days, zero when not overdue
    bValid : BOOL; // 结果有效位 [-] / result valid flag
    bOverdue : BOOL; // 逾期标志 [-] / overdue flag
    iErrCode : INT; // 事件码 0=正常 1=周期超域 2=上次时刻未初始化 3=秒计数溢出 / event code
END_VAR
VAR CONSTANT
    diSecPerDay : DINT := 86400; // 每日秒数 [s/d] / seconds per day
    diIntervalMax : DINT := 3650; // 周期天数上限 [d] / interval upper bound
END_VAR
VAR
    diLastSec : DINT; // 上次 PM 秒计数 [s] / last PM as seconds
    diNowSec : DINT; // 当前时刻秒计数 [s] / now as seconds
    diSpanSec : DINT; // 周期秒数 [s] / interval in seconds
    diNextSec : DINT; // 下次 PM 秒计数 [s] / next due as seconds
    diDiffSec : DINT; // 逾期秒数 [s] / overdue seconds
END_VAR

    // —— 段 0：全路径预清 —— //
    diLastSec := 0;
    diNowSec := 0;
    diSpanSec := 0;
    diNextSec := 0;
    diDiffSec := 0;
    dtNext := dtLast;
    dNextDate := DT_TO_DATE(dtLast);
    iOverdueDays := 0;
    bValid := FALSE;
    bOverdue := FALSE;
    iErrCode := 0;
    FC_DL_PmScheduleNext := FALSE;
    // —— 段 1：周期域闸 (0, 3650]d —— //
    IF (iIntervalDays <= 0) OR (INT_TO_DINT(iIntervalDays) > diIntervalMax) THEN
        iErrCode := 1; // 周期超域，不生成计划 / interval out of domain, no schedule issued
        RETURN;
    END_IF;
    // —— 段 2：上次时刻有效性闸（零值 = 未初始化） —— //
    diLastSec := DT_TO_DINT(dtLast); // 上次 PM 秒计数 [s] / last PM in seconds
    IF diLastSec <= 0 THEN
        iErrCode := 2; // 上次时刻未初始化 / last timestamp not initialised
        RETURN;
    END_IF;
    // —— 段 3：量纲链 (d)×(s/d) = s；加法后反查是否溢出为负 —— //
    diSpanSec := INT_TO_DINT(iIntervalDays) * diSecPerDay; // 周期秒数 [s] / interval in seconds
    diNextSec := diLastSec + diSpanSec; // 下次秒计数 [s] / next due in seconds
    IF diNextSec < diLastSec THEN
        iErrCode := 3; // 秒计数溢出，放弃本次计划 / second counter overflow, schedule dropped
        RETURN;
    END_IF;
    dtNext := DINT_TO_DT(diNextSec); // 下次到期时刻 [DT] / next due timestamp
    dNextDate := DT_TO_DATE(dtNext); // 到期日期 [DATE] / due date
    // —— 段 4：逾期天数 = MAX(0, (now-next)/86400) —— //
    diNowSec := DT_TO_DINT(dtNow); // 当前秒计数 [s] / now in seconds
    IF diNowSec > diNextSec THEN
        diDiffSec := diNowSec - diNextSec; // 逾期秒数 [s] / overdue seconds
        iOverdueDays := DINT_TO_INT(diDiffSec / diSecPerDay); // 逾期天数 [d] / overdue days
        bOverdue := TRUE;
    ELSE
        bOverdue := FALSE; // 未逾期 / not overdue
    END_IF;
    bValid := TRUE;
    FC_DL_PmScheduleNext := TRUE;
END_FUNCTION

(* ---- FC_DL_PneuAirConsumeCalc.st ---- *)
(*
  ============================================================
  组件名 : FC_DL_PneuAirConsumeCalc
  分类   : DL_Device
  功能   : 气缸耗气量计算，按缸径行程、表压与动作频次求单次与每分钟标准状态耗气量
  开源溯源 : internal-design（本轮无外部代码逐行引用）
             参考语义 : 无外部参考
  复杂度 : C1
  版本   : 1.0.0
  ============================================================
*)

FUNCTION FC_DL_PneuAirConsumeCalc : REAL
VAR_INPUT
    rBoreDia_mm    : REAL; // 缸径 [mm] bore diameter [mm]
    rStroke_mm     : REAL; // 行程 [mm] stroke [mm]
    rPressBar      : REAL; // 工作表压 [bar] working gauge pressure [bar]
    nCyclesPerMin  : INT; // 每分钟动作次数 [次/分] cycles per minute [cycle per minute]
    bDoubleActing  : BOOL; // 真为双作用，假为单作用 double acting when true, single acting when false
END_VAR
VAR_OUTPUT
    rAirPerCycle_Nl : REAL; // 单次耗气量（标准状态）[Nl] air per cycle at standard state [normal litre]
    rAirPerMin_Nl   : REAL; // 每分钟耗气量（标准状态）[Nl/min] air per minute at standard state [normal litre per minute]
    bValid          : BOOL; // 结果有效标志 result validity flag
END_VAR
VAR CONSTANT
    DL_PI_4      : REAL := 0.7853982; // 四分之圆周率 pi divided by four
    DL_MM3_PER_L : REAL := 1000000.0; // 每升立方毫米数 cubic millimetres per litre
    DL_ATM_BAR   : REAL := 1.013; // 标准大气压 [bar] standard atmosphere [bar]
    DL_TWO       : REAL := 2.0; // 双作用腔数因子 the double acting chamber factor
END_VAR
VAR
    _bFin  : BOOL := FALSE; // 三实数输入有限性判定 finiteness verdict of the three real inputs
    _rArea : REAL := 0.0; // 缸径截面面积 [mm2] bore section area [mm2]
    _rVolL : REAL := 0.0; // 单行程几何容积 [l] geometric volume per stroke [litre]
    _rStdL : REAL := 0.0; // 单次标准状态容积 [Nl] standard state volume per cycle [normal litre]
END_VAR

// 段 1｜出口预置 preset the exit
FC_DL_PneuAirConsumeCalc := 0.0; // 缺省返回零 default zero return
rAirPerCycle_Nl := 0.0; // 单次耗气预置零 air per cycle preset to zero
rAirPerMin_Nl := 0.0; // 分钟耗气预置零 air per minute preset to zero
bValid := FALSE; // 计算完成前不认结果 unusable before the calculation
// 段 2｜非有限闸 finiteness gate
_bFin := (rBoreDia_mm = rBoreDia_mm) AND (rStroke_mm = rStroke_mm) AND (rPressBar = rPressBar); // 三输入自反判定 self comparison of the three inputs
IF NOT _bFin THEN
    RETURN; // 非有限即无效 non finite means invalid
END_IF
// 段 3｜几何与频次闸 geometry and cycle gate
IF (rBoreDia_mm <= 0.0) OR (rStroke_mm < 0.0) OR (rPressBar < 0.0) THEN
    RETURN; // 几何或压力非法 an illegal geometry or pressure
END_IF
IF nCyclesPerMin < 0 THEN
    RETURN; // 负频次属配置非法 a negative cycle count is an illegal configuration
END_IF
// 段 4｜几何容积与双作用折算 geometric volume and the double acting factor
_rArea := DL_PI_4 * rBoreDia_mm * rBoreDia_mm; // 缸径截面面积 bore section area
_rVolL := _rArea * rStroke_mm / DL_MM3_PER_L; // 单行程几何容积 volume per stroke
IF bDoubleActing THEN
    _rVolL := _rVolL * DL_TWO; // 双作用按两腔估算，杆径影响按忽略处理 double acting counts both chambers with the rod ignored
END_IF
// 段 5｜标准状态折算与分钟耗气 standard state conversion and the minute consumption
_rStdL := _rVolL * (rPressBar + DL_ATM_BAR); // 表压折算到标准状态 gauge pressure converted to the standard state
rAirPerCycle_Nl := _rStdL; // 单次耗气落定 land the per cycle consumption
rAirPerMin_Nl := _rStdL * INT_TO_REAL(nCyclesPerMin); // 分钟耗气落定 land the per minute consumption
bValid := TRUE; // 结果可用 result usable
FC_DL_PneuAirConsumeCalc := rAirPerMin_Nl; // 函数返回分钟耗气 return the per minute consumption
END_FUNCTION

(* ---- FC_DL_PneuCvFlowCalc.st ---- *)
(*
  ============================================================
  组件名 : FC_DL_PneuCvFlowCalc
  分类   : DL_Device
  功能   : 气动元件 Cv 值流量估算，含临界压比判据与标准状态流量折算
  开源溯源 : internal-design（本轮无外部代码逐行引用）
             参考语义 : 无外部参考
  复杂度 : C1
  版本   : 1.0.0
  ============================================================
  口径说明 : 流量系数 0.865 属工程选型估算口径，压力取阀前绝对压力 [bar]，
             温度取开尔文，比重取相对空气值；输出直接为标准状态体积流量 [Nm3/h]。
             该式量纲一致，用于选型估算，精确定型须以厂商流量曲线复核。
*)

FUNCTION FC_DL_PneuCvFlowCalc : REAL
VAR_INPUT
    rCv           : REAL; // 流量系数 Cv [无量纲] flow coefficient Cv [dimensionless]
    rUpPressBarA  : REAL; // 阀前绝对压力 [bar abs] upstream absolute pressure [bar abs]
    rDownPressBarA: REAL; // 阀后绝对压力 [bar abs] downstream absolute pressure [bar abs]
    rTempC        : REAL; // 气体温度 [摄氏度] gas temperature [degree celsius]
    rGasSg        : REAL; // 相对空气比重 [无量纲] specific gravity relative to air [dimensionless]
END_VAR
VAR_OUTPUT
    rFlowNm3h : REAL; // 标准状态体积流量 [Nm3/h] normal volume flow [Nm3 per hour]
    rCritical : BOOL; // 临界流（阻塞流）标志 choked flow flag
    bValid    : BOOL; // 结果有效标志 result validity flag
END_VAR
VAR CONSTANT
    DL_CV_COEF   : REAL := 0.865; // 选型估算系数 sizing estimation coefficient
    DL_CRIT_RATIO: REAL := 0.528; // 空气临界压比 the critical air pressure ratio
    DL_KELVIN    : REAL := 273.15; // 摄氏到开尔文偏移 celsius to kelvin offset
    DL_EPS_R     : REAL := 1.0E-6; // 实数零判定阈值 real zero threshold
END_VAR
VAR
    _bFin  : BOOL := FALSE; // 五输入有限性判定 finiteness verdict of the five inputs
    _rTempK : REAL := 0.0; // 绝对温度 [K] absolute temperature [K]
    _rRatio : REAL := 0.0; // 压差比 pressure drop ratio [dimensionless]
    _rFlow : REAL := 0.0; // 流量中间量 [Nm3/h] intermediate flow [Nm3 per hour]
END_VAR

// 段 1｜出口预置 preset the exit
FC_DL_PneuCvFlowCalc := 0.0; // 缺省返回零 default zero return
rFlowNm3h := 0.0; // 流量预置零 flow preset to zero
rCritical := FALSE; // 临界标志预置假 critical flag preset false
bValid := FALSE; // 计算完成前不认结果 unusable before the calculation
// 段 2｜非有限闸 finiteness gate
_bFin := (rCv = rCv) AND (rUpPressBarA = rUpPressBarA) AND (rDownPressBarA = rDownPressBarA) AND (rTempC = rTempC) AND (rGasSg = rGasSg); // 五输入自反判定 self comparison of the five inputs
IF NOT _bFin THEN
    RETURN; // 非有限即无效 non finite means invalid
END_IF
// 段 3｜压力与介质闸 pressure and medium gate
IF (rUpPressBarA <= 0.0) OR (rDownPressBarA < 0.0) OR (rDownPressBarA > rUpPressBarA) THEN
    RETURN; // 阀前后压力倒置或非正 an inverted or non positive pressure pair
END_IF
IF (rGasSg <= 0.0) OR (rCv < 0.0) THEN
    RETURN; // 比重非正或 Cv 为负属配置非法 an illegal specific gravity or Cv
END_IF
// 段 4｜绝对温度与压差比 absolute temperature and the drop ratio
_rTempK := rTempC + DL_KELVIN; // 摄氏折算开尔文 convert celsius to kelvin
IF _rTempK <= DL_EPS_R THEN
    RETURN; // 绝对温度非正无法开方 a non positive absolute temperature cannot be rooted
END_IF
_rRatio := (rUpPressBarA - rDownPressBarA) / rUpPressBarA; // 压差比，除子已证为正 the drop ratio over a proven positive divisor
rCritical := _rRatio >= DL_CRIT_RATIO; // 达临界压比按阻塞流口径处理 a reached ratio is treated as choked flow
// 段 5｜主体流量估算 main flow estimation
_rFlow := DL_CV_COEF * rCv * rUpPressBarA * SQRT(1.0 / (rGasSg * _rTempK)); // 选型估算式，除子已证为正 the sizing formula over a proven positive divisor
rFlowNm3h := _rFlow; // 流量落定 land the flow
bValid := TRUE; // 结果可用 result usable
FC_DL_PneuCvFlowCalc := _rFlow; // 函数返回流量 return the flow
END_FUNCTION

(* ---- FC_DL_PneuLeakRateCalc.st ---- *)
(*
  ============================================================
  组件名 : FC_DL_PneuLeakRateCalc
  分类   : DL_Device
  功能   : 气密保压试验泄漏率计算，由起止压力、容积与试验时长求泄漏量与压降百分比
  开源溯源 : internal-design（本轮无外部代码逐行引用）
             参考语义 : 无外部参考
  复杂度 : C1
  版本   : 1.0.0
  ============================================================
*)

FUNCTION FC_DL_PneuLeakRateCalc : REAL
VAR_INPUT
    rPressStart_bar : REAL; // 试验起始压力 [bar] test start pressure [bar]
    rPressEnd_bar   : REAL; // 试验结束压力 [bar] test end pressure [bar]
    rVolume_l       : REAL; // 试件与管路容积 [l] specimen and piping volume [litre]
    rTestTimeS      : REAL; // 保压试验时长 [s] holding test duration [s]
    rTempC          : REAL; // 试验环境温度 [摄氏度] ambient test temperature [degree celsius]
END_VAR
VAR_OUTPUT
    rLeak_lpm      : REAL; // 标准状态泄漏量 [Nl/min] leak rate at standard state [normal litre per minute]
    rLeakPctPerMin : REAL; // 每分钟压降百分比 [%/min] pressure decay percentage per minute [% per minute]
    bValid         : BOOL; // 结果有效标志 result validity flag
END_VAR
VAR CONSTANT
    DL_ATM_BAR   : REAL := 1.01325; // 标准大气压 [bar] standard atmosphere [bar]
    DL_SEC_PER_MIN : REAL := 60.0; // 每分钟秒数 seconds per minute
    DL_KELVIN    : REAL := 273.15; // 摄氏到开尔文偏移 celsius to kelvin offset
    DL_T_REF_K   : REAL := 293.15; // 标准状态参考温度 [K] reference temperature at standard state [K]
    DL_HUNDRED   : REAL := 100.0; // 百分制换算系数 percentage scale factor
    DL_EPS_R     : REAL := 1.0E-6; // 实数零判定阈值 real zero threshold
END_VAR
VAR
    _bFin    : BOOL := FALSE; // 五输入有限性判定 finiteness verdict of the five inputs
    _rDropBar: REAL := 0.0; // 压力降 [bar] pressure drop [bar]
    _rTempK  : REAL := 0.0; // 绝对温度 [K] absolute temperature [K]
    _rVolStd : REAL := 0.0; // 标准状态泄漏体积 [Nl] normal leak volume [normal litre]
    _rLeak   : REAL := 0.0; // 泄漏量中间量 [Nl/min] intermediate leak rate [normal litre per minute]
    _rPct    : REAL := 0.0; // 每分钟压降百分比中间量 [%/min] intermediate decay percentage [% per minute]
END_VAR

// 段 1｜出口预置 preset the exit
FC_DL_PneuLeakRateCalc := 0.0; // 缺省返回零 default zero return
rLeak_lpm := 0.0; // 泄漏量预置零 leak rate preset to zero
rLeakPctPerMin := 0.0; // 压降百分比预置零 decay percentage preset to zero
bValid := FALSE; // 计算完成前不认结果 unusable before the calculation
// 段 2｜非有限闸 finiteness gate
_bFin := (rPressStart_bar = rPressStart_bar) AND (rPressEnd_bar = rPressEnd_bar) AND (rVolume_l = rVolume_l) AND (rTestTimeS = rTestTimeS) AND (rTempC = rTempC); // 五输入自反判定 self comparison of the five inputs
IF NOT _bFin THEN
    RETURN; // 非有限即无效 non finite means invalid
END_IF
// 段 3｜时长压力与容积闸 duration pressure and volume gate
IF (rTestTimeS <= DL_EPS_R) OR (rPressStart_bar <= DL_EPS_R) OR (rVolume_l <= 0.0) THEN
    RETURN; // 时长压力容积非正无法折算 a non positive duration pressure or volume cannot be converted
END_IF
IF rPressEnd_bar < 0.0 THEN
    RETURN; // 终压为负属采集异常 a negative end pressure is a measurement fault
END_IF
// 段 4｜标准状态泄漏体积 normal leak volume
_rDropBar := rPressStart_bar - rPressEnd_bar; // 试验段压力降 pressure drop over the test window
_rTempK := rTempC + DL_KELVIN; // 摄氏折算开尔文 convert celsius to kelvin
IF _rTempK <= DL_EPS_R THEN
    RETURN; // 绝对温度非正无法折算 a non positive absolute temperature cannot be converted
END_IF
_rVolStd := _rDropBar * rVolume_l / DL_ATM_BAR * (DL_T_REF_K / _rTempK); // 压降乘容积折标准状态 drop times volume normalised to the standard state
// 段 5｜泄漏率与压降百分比 leak rate and the decay percentage
_rLeak := _rVolStd / rTestTimeS * DL_SEC_PER_MIN; // 折算到每分钟 per minute leak rate
_rPct := (_rDropBar / rPressStart_bar * DL_HUNDRED) / (rTestTimeS / DL_SEC_PER_MIN); // 每分钟压降百分比 pressure decay percentage per minute
IF (_rLeak <> _rLeak) OR (ABS(_rLeak) > 1.0E30) OR (_rPct <> _rPct) OR (ABS(_rPct) > 1.0E30) THEN
    RETURN; // 结果非有限拒收 refuse a non finite result
END_IF
rLeak_lpm := _rLeak; // 泄漏量落定 land the leak rate
rLeakPctPerMin := _rPct; // 压降百分比落定 land the decay percentage
bValid := TRUE; // 结果可用 result usable
FC_DL_PneuLeakRateCalc := _rLeak; // 函数返回泄漏量 return the leak rate
END_FUNCTION

(* ---- FC_DL_PueInstantCalc.st ---- *)
(*
 * FC_DL_PueInstantCalc | C1 | DL_Device
 * 功能：瞬时 PUE 与 IT 负载占比       单位：功率 [kW]、PUE [1]、占比 [%]
 * 工况边界：仅适用于整机房口径（总功率含制冷、输配与照明，不小于 IT 功率）；IT 功率须 >0（入分母），否则判 9621；总功率小于 IT 功率说明计量口径错误，置 xValid=FALSE 但保留数值供诊断
 * 代数值回代：IT=500 kW、Total=700 kW → PUE=1.40、IT 占比 71.43 %（与 spec 回代行一致）
 * 开源溯源：clean-room 自研，未复制任何第三方代码（无外部来源）
 *)
FUNCTION FC_DL_PueInstantCalc : BOOL
VAR_INPUT
    rItKw    : REAL := 500.0;        // IT 设备功率 | IT equipment power [kW]
    rTotalKw : REAL := 700.0;        // 机房总功率 | total facility power [kW]
END_VAR
VAR_OUTPUT
    rPue      : REAL;                // 瞬时 PUE | instantaneous PUE [1]
    rItSharePct : REAL;              // IT 负载占比 | IT load share [%]
    xValid    : BOOL;                // 输出有效 | outputs valid
    nFaultCode: INT;                 // 0=无 / 9621=IT 功率非法 / 9622=总功率小于 IT 功率 | 0 none, 9621 illegal IT power, 9622 total below IT
END_VAR
VAR
    xFinIt : BOOL;                   // IT 功率有限性 | IT power is finite
    xFinTot: BOOL;                   // 总功率有限性 | total power is finite
END_VAR
VAR CONSTANT
    DL_PUE_PCT   : REAL := 100.0;    // 百分数换算系数 | percentage factor [%]
    DL_PUE_ITMIN : REAL := 1.0E-9;   // IT 功率下限（防零除）| IT power lower bound guarding the division [kW]
END_VAR

// 段1｜非有限闸（R19）
xFinIt := (rItKw = rItKw) AND ((rItKw - rItKw) = 0.0);
xFinTot := (rTotalKw = rTotalKw) AND ((rTotalKw - rTotalKw) = 0.0);
IF (NOT xFinIt) OR (NOT xFinTot) THEN
    rPue := 0.0;                     // 安全值：PUE 0（下游按无效丢弃）| safe value, downstream discards it
    rItSharePct := 0.0;
    xValid := FALSE;
    nFaultCode := 9621;
    FC_DL_PueInstantCalc := FALSE;
    RETURN;
END_IF

// 段2｜域闸：IT 功率入分母必须 >0，总功率不得为负
IF (rItKw <= DL_PUE_ITMIN) OR (rTotalKw < 0.0) THEN
    rPue := 0.0;
    rItSharePct := 0.0;
    xValid := FALSE;
    nFaultCode := 9621;
    FC_DL_PueInstantCalc := FALSE;
    RETURN;
END_IF

// 段3｜算法：PUE = 总功率/IT 功率；IT 占比同源
rPue := rTotalKw / rItKw;
rItSharePct := rItKw / rTotalKw * DL_PUE_PCT;

// 段4｜口径校验：总功率必须不小于 IT 功率（判据与出口同源于原始值）
IF rTotalKw < rItKw THEN
    xValid := FALSE;
    nFaultCode := 9622;              // 计量口径错误：数值保留供诊断，标志置无效 | metering inconsistency, value kept for diagnostics
    FC_DL_PueInstantCalc := FALSE;
    RETURN;
END_IF

// 段5｜出口
nFaultCode := 0;
xValid := TRUE;
FC_DL_PueInstantCalc := TRUE;
END_FUNCTION

(* ---- FC_DL_RackAirflowDemandCalc.st ---- *)
(*
 * FC_DL_RackAirflowDemandCalc | C2 | DL_Device
 * 功能：按机柜热负荷与允许温升反算所需送风量       单位：热负荷 [kW]、温升 [K]、密度 [kg/m³]、比热 [kJ/(kg·K)]、风量 [m³/h]
 * 工况边界：仅适用于封闭冷通道的机柜级风量估算（假定全部热负荷由送风带走，无旁通）；温升 rDeltaTC 须 >0（入分母），密度与比热须 >0；热负荷为 0 时风量为 0 仍有效
 * 代数值回代：Q=8 kW、ΔT=12 K、ρ=1.2、cp=1.005 → 3600×8/(1.2×1.005×12)=1990.0 m³/h（spec 记 1990 m³/h，一致）
 * 开源溯源：clean-room 自研，未复制任何第三方代码（无外部来源）
 *)
FUNCTION FC_DL_RackAirflowDemandCalc : BOOL
VAR_INPUT
    rRackLoadKw : REAL := 8.0;       // 机柜热负荷 | rack heat load [kW]
    rDeltaTC    : REAL := 12.0;      // 允许进回风温升 | permitted inlet to outlet temperature rise [K]
    rRho        : REAL := 1.2;       // 空气密度 | air density [kg/m³]
    rCp         : REAL := 1.005;     // 空气定压比热 | air specific heat at constant pressure [kJ/(kg·K)]
END_VAR
VAR_OUTPUT
    rAirflowM3h : REAL;              // 需求送风量 | required supply airflow [m³/h]
    xValid      : BOOL;              // 输出有效 | outputs valid
END_VAR
VAR
    xFinQ   : BOOL;                  // 热负荷有限性 | heat load is finite
    xFinDT  : BOOL;                  // 温升有限性 | temperature rise is finite
    xFinRho : BOOL;                  // 密度有限性 | density is finite
    xFinCp  : BOOL;                  // 比热有限性 | specific heat is finite
    rDen    : REAL;                  // 分母 ρ×cp×ΔT | denominator rho times cp times delta T [kW/(m³/h)]
END_VAR
VAR CONSTANT
    DL_RAD_SEC_PER_HOUR : REAL := 3600.0;  // 秒转小时系数 | seconds to hours factor [s/h]
    DL_RAD_DEN_MIN      : REAL := 1.0E-9;  // 除零保护阈值 | division guard threshold [kW/(m³/h)]
END_VAR

// 段1｜非有限闸（R19）
xFinQ := (rRackLoadKw = rRackLoadKw) AND ((rRackLoadKw - rRackLoadKw) = 0.0);
xFinDT := (rDeltaTC = rDeltaTC) AND ((rDeltaTC - rDeltaTC) = 0.0);
xFinRho := (rRho = rRho) AND ((rRho - rRho) = 0.0);
xFinCp := (rCp = rCp) AND ((rCp - rCp) = 0.0);
IF (NOT xFinQ) OR (NOT xFinDT) OR (NOT xFinRho) OR (NOT xFinCp) THEN
    rAirflowM3h := 0.0;              // 安全值：风量 0 | safe value, zero airflow
    xValid := FALSE;
    FC_DL_RackAirflowDemandCalc := FALSE;
    RETURN;
END_IF

// 段2｜域闸：温升入分母必须 >0，密度与比热须 >0，热负荷不得为负
IF (rDeltaTC <= 0.0) OR (rRho <= 0.0) OR (rCp <= 0.0) OR (rRackLoadKw < 0.0) THEN
    rAirflowM3h := 0.0;
    xValid := FALSE;
    FC_DL_RackAirflowDemandCalc := FALSE;
    RETURN;
END_IF

// 段3｜算法：V(m³/h) = 3600×Q/(ρ×cp×ΔT)，分母显式防零
rDen := rRho * rCp * rDeltaTC;
IF rDen > DL_RAD_DEN_MIN THEN
    rAirflowM3h := DL_RAD_SEC_PER_HOUR * rRackLoadKw / rDen;
ELSE
    rAirflowM3h := 0.0;              // 理论不可达（段2已排除），防御性兜底 | unreachable defence
END_IF

// 段4｜出口
xValid := TRUE;
FC_DL_RackAirflowDemandCalc := TRUE;
END_FUNCTION

(* ---- FC_DL_RawMealResidueCalc.st ---- *)
(*
  DL Factory R84 | FC_DL_RawMealResidueCalc
  功能：生料 80µm/200µm 双档筛余与细度系数，按目标带判合格并给磨机加减料建议
  开源溯源：无（clean-room 自研，依据公开工艺公式，来源=行业通用公式，许可证=MIT，借鉴点=公式结构）
  规则：R1-R16 全遵守
*)
FUNCTION FC_DL_RawMealResidueCalc : REAL
VAR_INPUT
    fRes80 : REAL := 14.0; // 80µm 筛余 [%] / residue on the 80 micron sieve [%]
    fRes200Um : REAL := 1.8; // 200µm 筛余实测值 [%] / residue on the 200 micron sieve [%]
    fLo80 : REAL := 10.0; // 80µm 筛余合格下限 [%] / lower acceptance bound [%]
    fHi80 : REAL := 18.0; // 80µm 筛余合格上限 [%] / upper acceptance bound [%]
END_VAR
VAR_OUTPUT
    fRes200 : REAL; // 200µm 筛余回显（链路校验） [%] / 200 micron residue echo [%]
    iAdvice : INT; // 磨机建议 1=加料 0=保持 −1=减料 [-] / mill advice [-]
    xPass : BOOL; // 细度判合格 [-] / fineness passed [-]
    xValid : BOOL; // 计算结果有效标志 [-] / calculation valid flag [-]
END_VAR
VAR
    fFinCoef : REAL; // 细度系数（80µm/200µm 比值） [-] / fineness coefficient [-]
END_VAR

// 段 1｜出口预置（R256）
FC_DL_RawMealResidueCalc := -1.0; // 哨兵返回 -1（无效） [-] / sentinel return -1, invalid [-]
fRes200 := 0.0; // 200µm 筛余回显预置零 [%] / residue echo preset zero [%]
iAdvice := 0; // 建议预置保持 [-] / advice preset to hold [-]
xPass := FALSE; // 合格位预置 FALSE [-] / pass preset false [-]
xValid := FALSE; // 计算完成前不认结果 [-] / unusable before calculation [-]

// 段 2｜非有限拦截 + 域闸（R4/R20）
IF NOT (fRes80 > -1.0E30 AND fRes80 < 1.0E30) OR NOT (fRes200Um > -1.0E30 AND fRes200Um < 1.0E30) OR NOT (fLo80 > -1.0E30 AND fLo80 < 1.0E30) OR NOT (fHi80 > -1.0E30 AND fHi80 < 1.0E30) THEN
    RETURN; // 任一入参为 NaN/Inf 一律拒绝 [-] / any NaN or Inf input rejected [-]
END_IF
IF fRes80 < 0.0 OR fRes200Um < 0.0 OR fRes80 > 100.0 OR fRes200Um > 100.0 THEN
    RETURN; // 筛余百分比域闸 (0~100) [%] / residue percentage domain gate [%]
END_IF
IF NOT (fLo80 < fHi80) THEN
    RETURN; // 目标带组态闸：下限必须严格小于上限 [%] / acceptance band config gate [%]
END_IF

// 段 3｜细度系数（200µm 筛余趋零时按极小值兜底）
fFinCoef := fRes80 / MAX(fRes200Um, 1.0E-9); // % ÷ % = 无量纲（比值越大即粗颗粒占比越集中） / [%] / [%] = [-]
IF NOT (fFinCoef > -1.0E30 AND fFinCoef < 1.0E30) THEN
    RETURN; // 结果非有限再拦一次 [-] / second finiteness gate [-]
END_IF

// 段 4｜合格判定与磨机建议（筛余偏高=偏粗→减料；偏低=偏细→加料）
IF fRes80 > fHi80 THEN
    iAdvice := -1; // 偏粗：建议减料（提高粉磨细度） [-] / coarse, reduce the feed [-]
    xPass := FALSE; // 超上限不合格 [-] / above the band, fail [-]
ELSIF fRes80 < fLo80 THEN
    iAdvice := 1; // 偏细：建议加料（提高产量） [-] / fine, increase the feed [-]
    xPass := FALSE; // 低于下限同样不合格（细度即电耗） [-] / below the band, fail [-]
ELSE
    iAdvice := 0; // 带内：保持当前喂料 [-] / in band, hold the feed [-]
    xPass := TRUE; // 带内合格 [-] / in band, pass [-]
END_IF
fRes200 := fRes200Um; // 回显 200µm 筛余实测值（校验链路量） [%] / echo the 200 micron residue [%]
xValid := TRUE; // 链路有效 [-] / chain valid [-]
FC_DL_RawMealResidueCalc := fRes80; // 返回 80µm 筛余 [%] / return the 80 micron residue [%]
END_FUNCTION

(* ---- FC_DL_RefCompressorCapacity.st ---- *)
(*
  ============================================================
  组件名 : FC_DL_RefCompressorCapacity
  分类   : DL_Device
  功能   : 压缩机质量流量与制冷量估算，按理论排量、转速比、容积效率与吸气密度折算
  开源溯源 : internal-design（本轮无外部代码逐行引用）
             参考语义 : 无外部参考
  复杂度 : C1
  版本   : 1.0.0
  ============================================================
*)

FUNCTION FC_DL_RefCompressorCapacity : REAL
VAR_INPUT
    rSweptVol_m3h    : REAL; // 理论排气量 [m3/h] theoretical swept volume [m3 per hour]
    rSpeed_rpm       : REAL; // 实测转速 [rpm] measured rotational speed [rpm]
    rSpeedRated_rpm  : REAL; // 额定转速 [rpm] rated rotational speed [rpm]
    rVolEff          : REAL; // 容积效率 0~1 [无量纲] volumetric efficiency from zero to one [dimensionless]
    rSuctionDens_kgm3: REAL; // 吸气密度 [kg/m3] suction gas density [kg per cubic metre]
    rDh_kJkg         : REAL; // 吸气到排气的焓差 [kJ/kg] enthalpy rise from suction to discharge [kJ per kilogram]
END_VAR
VAR_OUTPUT
    rMassFlow_kgh : REAL; // 质量流量 [kg/h] mass flow [kg per hour]
    rCapEst_kW    : REAL; // 估算制冷量 [kW] estimated cooling capacity [kW]
    bValid        : BOOL; // 结果有效标志 result validity flag
END_VAR
VAR CONSTANT
    DL_SEC_PER_HOUR : REAL := 3600.0; // 每小时秒数 seconds per hour
END_VAR
VAR
    _bFin  : BOOL := FALSE; // 六输入有限性判定 finiteness verdict of the six inputs
    _rSpeedRatio : REAL := 0.0; // 转速比 [无量纲] speed ratio [dimensionless]
    _rMass : REAL := 0.0; // 质量流量中间量 [kg/h] intermediate mass flow [kg per hour]
    _rCap  : REAL := 0.0; // 制冷量中间量 [kW] intermediate capacity [kW]
END_VAR

// 段 1｜出口预置 preset the exit
FC_DL_RefCompressorCapacity := 0.0; // 缺省返回零 default zero return
rMassFlow_kgh := 0.0; // 质量流量预置零 mass flow preset to zero
rCapEst_kW := 0.0; // 制冷量预置零 capacity preset to zero
bValid := FALSE; // 计算完成前不认结果 unusable before the calculation
// 段 2｜非有限闸 finiteness gate
_bFin := (rSweptVol_m3h = rSweptVol_m3h) AND (rSpeed_rpm = rSpeed_rpm) AND (rSpeedRated_rpm = rSpeedRated_rpm) AND (rVolEff = rVolEff) AND (rSuctionDens_kgm3 = rSuctionDens_kgm3) AND (rDh_kJkg = rDh_kJkg); // 六输入自反判定 self comparison of the six inputs
IF NOT _bFin THEN
    RETURN; // 非有限即无效 non finite means invalid
END_IF
// 段 3｜转速与效率闸 speed and efficiency gate
IF (rSpeedRated_rpm <= 0.0) OR (rSpeed_rpm < 0.0) THEN
    RETURN; // 额定转速非正或负转速 an illegal rated or measured speed
END_IF
IF (rVolEff <= 0.0) OR (rVolEff > 1.0) THEN
    RETURN; // 容积效率越出零到一 volumetric efficiency outside the open closed interval
END_IF
IF (rSweptVol_m3h < 0.0) OR (rSuctionDens_kgm3 <= 0.0) OR (rDh_kJkg <= 0.0) THEN
    RETURN; // 排量密度或焓差非法 an illegal swept volume density or enthalpy rise
END_IF
// 段 4｜转速比与质量流量 speed ratio and the mass flow
_rSpeedRatio := rSpeed_rpm / rSpeedRated_rpm; // 转速比，除子已证为正 speed ratio over a proven positive divisor
_rMass := rSweptVol_m3h * _rSpeedRatio * rVolEff * rSuctionDens_kgm3; // 排量乘转速比效率密度 swept volume times ratio efficiency and density
rMassFlow_kgh := _rMass; // 质量流量落定 land the mass flow
// 段 5｜焓差折算制冷量 enthalpy rise converted to capacity
_rCap := _rMass * rDh_kJkg / DL_SEC_PER_HOUR; // 千焦每小时折算为千瓦 kilojoule per hour becomes kilowatt
rCapEst_kW := _rCap; // 制冷量落定 land the capacity
bValid := TRUE; // 结果可用 result usable
FC_DL_RefCompressorCapacity := _rMass; // 函数返回质量流量 return the mass flow
END_FUNCTION

(* ---- FC_DL_RefCondApproach.st ---- *)
(*
  ============================================================
  组件名 : FC_DL_RefCondApproach
  分类   : DL_Device
  功能   : 冷凝器逼近度计算，由冷凝饱和温度与进风温度求逼近度并判换热面污染
  开源溯源 : internal-design（本轮无外部代码逐行引用）
             参考语义 : 无外部参考
  复杂度 : C1
  版本   : 1.0.0
  ============================================================
*)

FUNCTION FC_DL_RefCondApproach : REAL
VAR_INPUT
    rCondSatTempC   : REAL; // 冷凝饱和温度 [摄氏度] condensing saturation temperature [degree celsius]
    rAirInTempC     : REAL; // 冷凝器进风温度 [摄氏度] condenser entering air temperature [degree celsius]
    rApproachRef    : REAL; // 设计逼近度基准 [K] design approach reference [kelvin]
    rApproachAlarm  : REAL; // 逼近度报警限 [K] approach alarm limit [kelvin]
END_VAR
VAR_OUTPUT
    rApproachK : REAL; // 实测逼近度 [K] measured approach [kelvin]
    bFouling   : BOOL; // 换热面污染判据标志 fouling verdict flag
    bValid     : BOOL; // 结果有效标志 result validity flag
END_VAR
VAR
    _bFin : BOOL := FALSE; // 四输入有限性判定 finiteness verdict of the four inputs
    _rAp  : REAL := 0.0; // 逼近度中间量 [K] intermediate approach [kelvin]
    _rLim : REAL := 0.0; // 钳位后的报警限 [K] clamped alarm limit [kelvin]
END_VAR

// 段 1｜出口预置 preset the exit
FC_DL_RefCondApproach := 0.0; // 缺省返回零 default zero return
rApproachK := 0.0; // 逼近度预置零 approach preset to zero
bFouling := FALSE; // 污染标志预置假 fouling flag preset false
bValid := FALSE; // 计算完成前不认结果 unusable before the calculation
// 段 2｜非有限闸 finiteness gate
_bFin := (rCondSatTempC = rCondSatTempC) AND (rAirInTempC = rAirInTempC) AND (rApproachRef = rApproachRef) AND (rApproachAlarm = rApproachAlarm); // 四输入自反判定 self comparison of the four inputs
IF NOT _bFin THEN
    RETURN; // 非有限即无效 non finite means invalid
END_IF
// 段 3｜主体逼近度 main approach
_rAp := rCondSatTempC - rAirInTempC; // 冷凝饱和温度减进风温度 condensing saturation minus the entering air
rApproachK := _rAp; // 逼近度落定 land the approach
// 段 4｜报警限整形与污染判定 alarm limit reshape and the fouling verdict
_rLim := rApproachAlarm; // 取入参报警限 take the alarm limit input
IF _rLim < 0.0 THEN
    _rLim := ABS(_rLim); // 负报警限取幅值 a negative limit becomes its magnitude
END_IF
bFouling := _rAp > _rLim; // 超限判换热面污染 an exceeded limit indicates fouling
bValid := TRUE; // 结果可用 result usable
FC_DL_RefCondApproach := _rAp; // 函数返回逼近度 return the approach
END_FUNCTION

(* ---- FC_DL_RefCopCalc.st ---- *)
(*
  ============================================================
  组件名 : FC_DL_RefCopCalc
  分类   : DL_Device
  功能   : 制冷机组能效比计算，由制冷量与输入功率求 COP 及其与额定值的比值
  开源溯源 : internal-design（本轮无外部代码逐行引用）
             参考语义 : 无外部参考
  复杂度 : C1
  版本   : 1.0.0
  ============================================================
*)

FUNCTION FC_DL_RefCopCalc : REAL
VAR_INPUT
    rCoolingCap_kW : REAL; // 制冷量 [kW] cooling capacity [kW]
    rPowerIn_kW    : REAL; // 输入功率 [kW] electrical power input [kW]
    rCopRated      : REAL; // 额定能效比 [无量纲] rated coefficient of performance [dimensionless]
END_VAR
VAR_OUTPUT
    rCop      : REAL; // 实测能效比 [无量纲] measured coefficient of performance [dimensionless]
    rCopRatio : REAL; // 实测与额定能效比之比 [无量纲] ratio of the measured to the rated value [dimensionless]
    bValid    : BOOL; // 结果有效标志 result validity flag
END_VAR
VAR CONSTANT
    DL_POWER_FLOOR : REAL := 0.01; // 功率有效下限 [kW] power effective floor [kW]
END_VAR
VAR
    _bFin  : BOOL := FALSE; // 三输入有限性判定 finiteness verdict of the three inputs
    _rCop  : REAL := 0.0; // 能效比中间量 [无量纲] intermediate coefficient [dimensionless]
    _rRat  : REAL := 0.0; // 比值中间量 [无量纲] intermediate ratio [dimensionless]
END_VAR

// 段 1｜出口预置 preset the exit
FC_DL_RefCopCalc := 0.0; // 缺省返回零 default zero return
rCop := 0.0; // 能效比预置零 coefficient preset to zero
rCopRatio := 0.0; // 比值预置零 ratio preset to zero
bValid := FALSE; // 计算完成前不认结果 unusable before the calculation
// 段 2｜非有限闸 finiteness gate
_bFin := (rCoolingCap_kW = rCoolingCap_kW) AND (rPowerIn_kW = rPowerIn_kW) AND (rCopRated = rCopRated); // 三输入自反判定 self comparison of the three inputs
IF NOT _bFin THEN
    RETURN; // 非有限即无效 non finite means invalid
END_IF
// 段 3｜功率分母闸 power divisor gate
IF rPowerIn_kW <= DL_POWER_FLOOR THEN
    RETURN; // 功率低于有效下限判无效 a power below the floor is void
END_IF
// 段 4｜主体能效比 main coefficient of performance
_rCop := rCoolingCap_kW / rPowerIn_kW; // 制冷量除以输入功率 capacity over the power input
rCop := _rCop; // 能效比落定 land the coefficient
// 段 5｜额定比值闸 rated ratio gate
IF rCopRated <= 0.0 THEN
    RETURN; // 额定值非正无法求比值 a non positive rating cannot carry a ratio
END_IF
_rRat := _rCop / rCopRated; // 实测对额定比值 measured over rated
rCopRatio := _rRat; // 比值落定 land the ratio
bValid := TRUE; // 结果可用 result usable
FC_DL_RefCopCalc := _rCop; // 函数返回能效比 return the coefficient
END_FUNCTION
